// --- Siemens Structured Format ---
DATA_BLOCK "model__HS32_IW10_"
{ S7_Optimized_Access := 'TRUE' }
VERSION :
NON_RETAIN
   VAR
      W_i : ARRAY[0..31, 0..39] OF REAL;
      W_f : ARRAY[0..31, 0..39] OF REAL;
      W_g : ARRAY[0..31, 0..39] OF REAL;
      W_o : ARRAY[0..31, 0..39] OF REAL;
      R_i : ARRAY[0..31, 0..31] OF REAL;
      R_f : ARRAY[0..31, 0..31] OF REAL;
      R_g : ARRAY[0..31, 0..31] OF REAL;
      R_o : ARRAY[0..31, 0..31] OF REAL;
      B_i : ARRAY[0..31] OF REAL;
      B_f : ARRAY[0..31] OF REAL;
      B_g : ARRAY[0..31] OF REAL;
      B_o : ARRAY[0..31] OF REAL;
      FC_W : ARRAY[0..39, 0..31] OF REAL;
      FC_B : ARRAY[0..39] OF REAL;
   END_VAR
BEGIN

      W_i[0,0] := -0.10414906;
      W_i[0,1] := 0.05087908;
      W_i[0,2] := 0.03123917;
      W_i[0,3] := 0.07883381;
      W_i[0,4] := -0.04182333;
      W_i[0,5] := -0.00272775;
      W_i[0,6] := -0.10306227;
      W_i[0,7] := 0.27651954;
      W_i[0,8] := 0.07111089;
      W_i[0,9] := -0.17811616;
      W_i[0,10] := 0.00811404;
      W_i[0,11] := 0.09247471;
      W_i[0,12] := -0.06765226;
      W_i[0,13] := 0.00099094;
      W_i[0,14] := -0.00565724;
      W_i[0,15] := 0.07034151;
      W_i[0,16] := -0.03319963;
      W_i[0,17] := -0.01640407;
      W_i[0,18] := 0.00714720;
      W_i[0,19] := 0.05200255;
      W_i[0,20] := -0.10294636;
      W_i[0,21] := 0.13340643;
      W_i[0,22] := -0.48219806;
      W_i[0,23] := -0.10634176;
      W_i[0,24] := -0.78127921;
      W_i[0,25] := -0.72295207;
      W_i[0,26] := -0.21058698;
      W_i[0,27] := -0.23595250;
      W_i[0,28] := -0.07997044;
      W_i[0,29] := -0.01075801;
      W_i[0,30] := -0.32065672;
      W_i[0,31] := -0.08546381;
      W_i[0,32] := -0.13408948;
      W_i[0,33] := 0.01877546;
      W_i[0,34] := -0.84940672;
      W_i[0,35] := -0.07448237;
      W_i[0,36] := -0.02454676;
      W_i[0,37] := -0.26921397;
      W_i[0,38] := -0.07333633;
      W_i[0,39] := -0.01266416;
      W_i[1,0] := 0.29037470;
      W_i[1,1] := 0.04892659;
      W_i[1,2] := 0.02171497;
      W_i[1,3] := 0.02552549;
      W_i[1,4] := 0.01215333;
      W_i[1,5] := 0.03346634;
      W_i[1,6] := -0.03770757;
      W_i[1,7] := 0.26558429;
      W_i[1,8] := -0.11029382;
      W_i[1,9] := -0.20845115;
      W_i[1,10] := -0.01400178;
      W_i[1,11] := 0.15223934;
      W_i[1,12] := -0.13050519;
      W_i[1,13] := -0.04419332;
      W_i[1,14] := 0.00628915;
      W_i[1,15] := 0.04288426;
      W_i[1,16] := -0.00701924;
      W_i[1,17] := 0.02646778;
      W_i[1,18] := -0.00136598;
      W_i[1,19] := 0.07391773;
      W_i[1,20] := 0.03997133;
      W_i[1,21] := 0.11501998;
      W_i[1,22] := -0.30713096;
      W_i[1,23] := -0.01738190;
      W_i[1,24] := -0.39384720;
      W_i[1,25] := -0.48897827;
      W_i[1,26] := -0.01727662;
      W_i[1,27] := -0.21526198;
      W_i[1,28] := -0.00675165;
      W_i[1,29] := 0.18086264;
      W_i[1,30] := -0.21994361;
      W_i[1,31] := -0.03053124;
      W_i[1,32] := -0.17159809;
      W_i[1,33] := -0.00609811;
      W_i[1,34] := -0.71118248;
      W_i[1,35] := -0.12901427;
      W_i[1,36] := -0.05088318;
      W_i[1,37] := -0.12064310;
      W_i[1,38] := -0.03252085;
      W_i[1,39] := -0.03171032;
      W_i[2,0] := -0.00230766;
      W_i[2,1] := -0.01114088;
      W_i[2,2] := 0.00278754;
      W_i[2,3] := -0.04560725;
      W_i[2,4] := -0.00076747;
      W_i[2,5] := -0.02340589;
      W_i[2,6] := -0.09104784;
      W_i[2,7] := -0.03890763;
      W_i[2,8] := 0.02353094;
      W_i[2,9] := 0.00039863;
      W_i[2,10] := 0.01153927;
      W_i[2,11] := 0.04803184;
      W_i[2,12] := 0.08744484;
      W_i[2,13] := 0.04118077;
      W_i[2,14] := 0.02094036;
      W_i[2,15] := 0.12591685;
      W_i[2,16] := 0.01395341;
      W_i[2,17] := 0.02091648;
      W_i[2,18] := -0.04870405;
      W_i[2,19] := -0.04149374;
      W_i[2,20] := 0.10584776;
      W_i[2,21] := 0.06836145;
      W_i[2,22] := 0.01589410;
      W_i[2,23] := -0.06229543;
      W_i[2,24] := -0.27194241;
      W_i[2,25] := -0.39684960;
      W_i[2,26] := 0.03680405;
      W_i[2,27] := 0.08170957;
      W_i[2,28] := 0.08198555;
      W_i[2,29] := 0.08877461;
      W_i[2,30] := 0.25039282;
      W_i[2,31] := 0.00393842;
      W_i[2,32] := 0.15045230;
      W_i[2,33] := -0.04096574;
      W_i[2,34] := 0.44737267;
      W_i[2,35] := -0.14432395;
      W_i[2,36] := -0.04863369;
      W_i[2,37] := -0.42030501;
      W_i[2,38] := -0.05893779;
      W_i[2,39] := -0.01147668;
      W_i[3,0] := -0.11661218;
      W_i[3,1] := -0.11039881;
      W_i[3,2] := -0.09505490;
      W_i[3,3] := -0.05274161;
      W_i[3,4] := 0.13631159;
      W_i[3,5] := -0.41682443;
      W_i[3,6] := 0.34413198;
      W_i[3,7] := 0.19693865;
      W_i[3,8] := -0.37381542;
      W_i[3,9] := 0.03602328;
      W_i[3,10] := 0.32276613;
      W_i[3,11] := -0.61351973;
      W_i[3,12] := -0.15591657;
      W_i[3,13] := -0.22586936;
      W_i[3,14] := -0.00271499;
      W_i[3,15] := 0.03598518;
      W_i[3,16] := -0.04658272;
      W_i[3,17] := 0.12849101;
      W_i[3,18] := 0.14830461;
      W_i[3,19] := 0.61608970;
      W_i[3,20] := -0.01793281;
      W_i[3,21] := 0.22755618;
      W_i[3,22] := 0.04441701;
      W_i[3,23] := 0.06841668;
      W_i[3,24] := -0.42572534;
      W_i[3,25] := -0.38698140;
      W_i[3,26] := 0.11054352;
      W_i[3,27] := -0.20471475;
      W_i[3,28] := -0.03201612;
      W_i[3,29] := -0.26479176;
      W_i[3,30] := 0.02552174;
      W_i[3,31] := -0.13836773;
      W_i[3,32] := -0.11162268;
      W_i[3,33] := -0.09296755;
      W_i[3,34] := -0.26265231;
      W_i[3,35] := -0.16597824;
      W_i[3,36] := 0.03927263;
      W_i[3,37] := -0.06124702;
      W_i[3,38] := 0.16334522;
      W_i[3,39] := 0.95440286;
      W_i[4,0] := -0.09592919;
      W_i[4,1] := 0.07784065;
      W_i[4,2] := 0.01346385;
      W_i[4,3] := 0.08287931;
      W_i[4,4] := -0.42782676;
      W_i[4,5] := 0.03361791;
      W_i[4,6] := -0.15880656;
      W_i[4,7] := -0.05813188;
      W_i[4,8] := -0.01824343;
      W_i[4,9] := -0.11751872;
      W_i[4,10] := 0.14676669;
      W_i[4,11] := 0.02209505;
      W_i[4,12] := -0.00572815;
      W_i[4,13] := 0.05958780;
      W_i[4,14] := -0.02038914;
      W_i[4,15] := -0.01525941;
      W_i[4,16] := -0.03268129;
      W_i[4,17] := 0.01159987;
      W_i[4,18] := -0.02004867;
      W_i[4,19] := -0.07593681;
      W_i[4,20] := 0.05724435;
      W_i[4,21] := -0.28372633;
      W_i[4,22] := -0.11699247;
      W_i[4,23] := -0.35998097;
      W_i[4,24] := 0.26990792;
      W_i[4,25] := 0.15219623;
      W_i[4,26] := -0.08656731;
      W_i[4,27] := 0.16333446;
      W_i[4,28] := 0.13229539;
      W_i[4,29] := 0.18428297;
      W_i[4,30] := -0.18249886;
      W_i[4,31] := 0.24244712;
      W_i[4,32] := -0.00069160;
      W_i[4,33] := 0.29610279;
      W_i[4,34] := 0.03106182;
      W_i[4,35] := -0.07256878;
      W_i[4,36] := 0.03714421;
      W_i[4,37] := -0.08504521;
      W_i[4,38] := -0.01051908;
      W_i[4,39] := 0.00350483;
      W_i[5,0] := -0.05495714;
      W_i[5,1] := 0.17977138;
      W_i[5,2] := 0.04651625;
      W_i[5,3] := 0.08715992;
      W_i[5,4] := 0.10765444;
      W_i[5,5] := -0.10662776;
      W_i[5,6] := -0.04317707;
      W_i[5,7] := 0.04963618;
      W_i[5,8] := 0.00394473;
      W_i[5,9] := 0.02992170;
      W_i[5,10] := -0.02726821;
      W_i[5,11] := 0.21677773;
      W_i[5,12] := -0.15348147;
      W_i[5,13] := -0.01556183;
      W_i[5,14] := 0.01471778;
      W_i[5,15] := -0.00319904;
      W_i[5,16] := 0.06557427;
      W_i[5,17] := -0.00420085;
      W_i[5,18] := 0.00420561;
      W_i[5,19] := 0.07868493;
      W_i[5,20] := -0.17903206;
      W_i[5,21] := -0.01610633;
      W_i[5,22] := -0.42383689;
      W_i[5,23] := -0.00551023;
      W_i[5,24] := -0.38271463;
      W_i[5,25] := -0.08532900;
      W_i[5,26] := 0.03424337;
      W_i[5,27] := 0.00513940;
      W_i[5,28] := -0.12665990;
      W_i[5,29] := 0.72981369;
      W_i[5,30] := -0.61144358;
      W_i[5,31] := -0.02451378;
      W_i[5,32] := -0.15765238;
      W_i[5,33] := -0.08363440;
      W_i[5,34] := -0.17316997;
      W_i[5,35] := 0.04921770;
      W_i[5,36] := 0.03656118;
      W_i[5,37] := -0.23534429;
      W_i[5,38] := -0.03259736;
      W_i[5,39] := -0.02564295;
      W_i[6,0] := -0.07149911;
      W_i[6,1] := 0.05910936;
      W_i[6,2] := 0.02579894;
      W_i[6,3] := 0.07767012;
      W_i[6,4] := -0.02382352;
      W_i[6,5] := 0.03319338;
      W_i[6,6] := -0.03900349;
      W_i[6,7] := -0.11483924;
      W_i[6,8] := -0.07984669;
      W_i[6,9] := -0.03000957;
      W_i[6,10] := 0.04087067;
      W_i[6,11] := 0.05389729;
      W_i[6,12] := -0.15653324;
      W_i[6,13] := -0.03200754;
      W_i[6,14] := -0.00524681;
      W_i[6,15] := -0.00143958;
      W_i[6,16] := -0.01686914;
      W_i[6,17] := -0.00267206;
      W_i[6,18] := 0.03467545;
      W_i[6,19] := 0.11881366;
      W_i[6,20] := 0.15485220;
      W_i[6,21] := -0.25145912;
      W_i[6,22] := 0.02979270;
      W_i[6,23] := 0.04974350;
      W_i[6,24] := -0.06280798;
      W_i[6,25] := 0.04208164;
      W_i[6,26] := 0.06788322;
      W_i[6,27] := 0.22705127;
      W_i[6,28] := 0.07820445;
      W_i[6,29] := -0.25283822;
      W_i[6,30] := 0.02389662;
      W_i[6,31] := -0.03982587;
      W_i[6,32] := 0.08894450;
      W_i[6,33] := 0.11913013;
      W_i[6,34] := 0.21554954;
      W_i[6,35] := -0.32464555;
      W_i[6,36] := 0.02452838;
      W_i[6,37] := -0.31377190;
      W_i[6,38] := 0.00847345;
      W_i[6,39] := 0.09918413;
      W_i[7,0] := 0.02757634;
      W_i[7,1] := -0.02689262;
      W_i[7,2] := -0.02939863;
      W_i[7,3] := -0.04568179;
      W_i[7,4] := -0.09635723;
      W_i[7,5] := -0.03179899;
      W_i[7,6] := -0.12191572;
      W_i[7,7] := 0.30427256;
      W_i[7,8] := 0.21273117;
      W_i[7,9] := -0.31949016;
      W_i[7,10] := 0.01761072;
      W_i[7,11] := -0.09866854;
      W_i[7,12] := 0.10523087;
      W_i[7,13] := 0.07799035;
      W_i[7,14] := 0.07163531;
      W_i[7,15] := 0.04057769;
      W_i[7,16] := -0.03791607;
      W_i[7,17] := 0.04264954;
      W_i[7,18] := -0.09266370;
      W_i[7,19] := -0.00260587;
      W_i[7,20] := -0.03977212;
      W_i[7,21] := -0.20910311;
      W_i[7,22] := -0.00171320;
      W_i[7,23] := -0.04438376;
      W_i[7,24] := -1.20630348;
      W_i[7,25] := -0.21321478;
      W_i[7,26] := -0.06407063;
      W_i[7,27] := 0.11449858;
      W_i[7,28] := 0.03520356;
      W_i[7,29] := 0.21331252;
      W_i[7,30] := 0.21956272;
      W_i[7,31] := -0.00092769;
      W_i[7,32] := -0.11663342;
      W_i[7,33] := 0.14221379;
      W_i[7,34] := -0.10930648;
      W_i[7,35] := 0.04132334;
      W_i[7,36] := 0.05281549;
      W_i[7,37] := 0.15278573;
      W_i[7,38] := 0.15391673;
      W_i[7,39] := -0.02757900;
      W_i[8,0] := 0.05724476;
      W_i[8,1] := -0.03158160;
      W_i[8,2] := -0.11627535;
      W_i[8,3] := -0.05773278;
      W_i[8,4] := 0.07278191;
      W_i[8,5] := -0.08000189;
      W_i[8,6] := 0.02300551;
      W_i[8,7] := -0.08800174;
      W_i[8,8] := 0.20740731;
      W_i[8,9] := 0.06626759;
      W_i[8,10] := 0.04762848;
      W_i[8,11] := -0.10821844;
      W_i[8,12] := -0.12422320;
      W_i[8,13] := 0.02703045;
      W_i[8,14] := 0.00398667;
      W_i[8,15] := 0.00804039;
      W_i[8,16] := -0.14637028;
      W_i[8,17] := -0.07778820;
      W_i[8,18] := -0.09220842;
      W_i[8,19] := 0.47469196;
      W_i[8,20] := 0.02264124;
      W_i[8,21] := 0.04296339;
      W_i[8,22] := 0.04171297;
      W_i[8,23] := -0.06263759;
      W_i[8,24] := 0.27121377;
      W_i[8,25] := 0.31945908;
      W_i[8,26] := 0.14077963;
      W_i[8,27] := 0.10558233;
      W_i[8,28] := -0.00015772;
      W_i[8,29] := 0.18647811;
      W_i[8,30] := 0.11800971;
      W_i[8,31] := 0.10110309;
      W_i[8,32] := 0.01555773;
      W_i[8,33] := 0.06486533;
      W_i[8,34] := 0.31461737;
      W_i[8,35] := 0.15680584;
      W_i[8,36] := -0.01419803;
      W_i[8,37] := 0.05979521;
      W_i[8,38] := 0.22562319;
      W_i[8,39] := 0.54453236;
      W_i[9,0] := -0.45409659;
      W_i[9,1] := -0.06150096;
      W_i[9,2] := 0.49318254;
      W_i[9,3] := -0.51527238;
      W_i[9,4] := 0.12728609;
      W_i[9,5] := -0.10118011;
      W_i[9,6] := 0.29715037;
      W_i[9,7] := -0.05259424;
      W_i[9,8] := 0.01368861;
      W_i[9,9] := 0.17207454;
      W_i[9,10] := 0.11617907;
      W_i[9,11] := 0.01172454;
      W_i[9,12] := -0.30126482;
      W_i[9,13] := 0.17993747;
      W_i[9,14] := 0.08894411;
      W_i[9,15] := -0.23540320;
      W_i[9,16] := -0.15334457;
      W_i[9,17] := -0.18120950;
      W_i[9,18] := 0.09745281;
      W_i[9,19] := 0.18141954;
      W_i[9,20] := 0.10671264;
      W_i[9,21] := 0.24788895;
      W_i[9,22] := 0.13593909;
      W_i[9,23] := -0.13985786;
      W_i[9,24] := -0.24154125;
      W_i[9,25] := -0.12681547;
      W_i[9,26] := 0.20098042;
      W_i[9,27] := -0.32428232;
      W_i[9,28] := -0.32814661;
      W_i[9,29] := -0.23453857;
      W_i[9,30] := 0.12634908;
      W_i[9,31] := 0.14591648;
      W_i[9,32] := -0.03520398;
      W_i[9,33] := 0.11785780;
      W_i[9,34] := -1.13588667;
      W_i[9,35] := -0.19602355;
      W_i[9,36] := 0.09494327;
      W_i[9,37] := 0.00611658;
      W_i[9,38] := 0.19538435;
      W_i[9,39] := 0.03790567;
      W_i[10,0] := 0.08093075;
      W_i[10,1] := -0.03189079;
      W_i[10,2] := 0.00460666;
      W_i[10,3] := -0.25079808;
      W_i[10,4] := 0.12079003;
      W_i[10,5] := 0.06994910;
      W_i[10,6] := 0.01222384;
      W_i[10,7] := 0.07541763;
      W_i[10,8] := 0.05855694;
      W_i[10,9] := -0.01396475;
      W_i[10,10] := 0.02662643;
      W_i[10,11] := -0.66687572;
      W_i[10,12] := 0.49504700;
      W_i[10,13] := -0.05885675;
      W_i[10,14] := -0.11757897;
      W_i[10,15] := 0.06344132;
      W_i[10,16] := -0.02143165;
      W_i[10,17] := 0.02022251;
      W_i[10,18] := -0.03556326;
      W_i[10,19] := 0.04088999;
      W_i[10,20] := -0.08695306;
      W_i[10,21] := 0.13901219;
      W_i[10,22] := -0.04673401;
      W_i[10,23] := -0.13039219;
      W_i[10,24] := -0.02369194;
      W_i[10,25] := -0.13022855;
      W_i[10,26] := 0.15325138;
      W_i[10,27] := -0.14148274;
      W_i[10,28] := -0.10921547;
      W_i[10,29] := 0.50673056;
      W_i[10,30] := 0.16923237;
      W_i[10,31] := -0.06320494;
      W_i[10,32] := -0.08798328;
      W_i[10,33] := 0.01157838;
      W_i[10,34] := -0.41323879;
      W_i[10,35] := 0.09598303;
      W_i[10,36] := 0.02359625;
      W_i[10,37] := -0.05013705;
      W_i[10,38] := -0.02053811;
      W_i[10,39] := 1.16537046;
      W_i[11,0] := -0.13920400;
      W_i[11,1] := 0.10422801;
      W_i[11,2] := 0.05192634;
      W_i[11,3] := 0.02474182;
      W_i[11,4] := -0.11992953;
      W_i[11,5] := -0.11497844;
      W_i[11,6] := -0.06959671;
      W_i[11,7] := 0.08906282;
      W_i[11,8] := 0.00035152;
      W_i[11,9] := -0.10795452;
      W_i[11,10] := 0.02394083;
      W_i[11,11] := -0.07669503;
      W_i[11,12] := 0.15492713;
      W_i[11,13] := 0.02082890;
      W_i[11,14] := 0.01739825;
      W_i[11,15] := 0.28620026;
      W_i[11,16] := -0.05672961;
      W_i[11,17] := 0.07933230;
      W_i[11,18] := -0.19136667;
      W_i[11,19] := -0.39791319;
      W_i[11,20] := -0.13187614;
      W_i[11,21] := -0.04277104;
      W_i[11,22] := -0.11175538;
      W_i[11,23] := -0.10681376;
      W_i[11,24] := -0.71706533;
      W_i[11,25] := -0.89369446;
      W_i[11,26] := -0.04355099;
      W_i[11,27] := -0.11690557;
      W_i[11,28] := 0.17073342;
      W_i[11,29] := 0.26696113;
      W_i[11,30] := -0.03069729;
      W_i[11,31] := -0.11184800;
      W_i[11,32] := 0.15421732;
      W_i[11,33] := 0.14543033;
      W_i[11,34] := -0.00053378;
      W_i[11,35] := 0.08841224;
      W_i[11,36] := 0.00902623;
      W_i[11,37] := -0.14363292;
      W_i[11,38] := -0.02996587;
      W_i[11,39] := 0.03438438;
      W_i[12,0] := 0.02294069;
      W_i[12,1] := -0.00171102;
      W_i[12,2] := -0.00742173;
      W_i[12,3] := -0.06263760;
      W_i[12,4] := 0.01279054;
      W_i[12,5] := -0.07051820;
      W_i[12,6] := 0.03081366;
      W_i[12,7] := 0.01733820;
      W_i[12,8] := -0.01632435;
      W_i[12,9] := -0.03842505;
      W_i[12,10] := 0.11362740;
      W_i[12,11] := 0.01187946;
      W_i[12,12] := -0.19036539;
      W_i[12,13] := 0.00812287;
      W_i[12,14] := 0.00857556;
      W_i[12,15] := 0.06468427;
      W_i[12,16] := 0.01327470;
      W_i[12,17] := 0.05196055;
      W_i[12,18] := 0.00679103;
      W_i[12,19] := 0.10192532;
      W_i[12,20] := 0.01617677;
      W_i[12,21] := -0.01601717;
      W_i[12,22] := -0.22829570;
      W_i[12,23] := 0.02394662;
      W_i[12,24] := -0.15263872;
      W_i[12,25] := -0.21143152;
      W_i[12,26] := 0.02614386;
      W_i[12,27] := 0.03263390;
      W_i[12,28] := -0.02625607;
      W_i[12,29] := 0.11965574;
      W_i[12,30] := -0.15762709;
      W_i[12,31] := -0.02538990;
      W_i[12,32] := -0.08307584;
      W_i[12,33] := -0.31617489;
      W_i[12,34] := -0.47193074;
      W_i[12,35] := 0.05056112;
      W_i[12,36] := -0.02334138;
      W_i[12,37] := 0.05162949;
      W_i[12,38] := -0.00184243;
      W_i[12,39] := -0.07476960;
      W_i[13,0] := -0.05422729;
      W_i[13,1] := 0.05369066;
      W_i[13,2] := 0.19673365;
      W_i[13,3] := -0.01662629;
      W_i[13,4] := -0.25112736;
      W_i[13,5] := 0.04215603;
      W_i[13,6] := -0.01216646;
      W_i[13,7] := -0.02261561;
      W_i[13,8] := 0.06583825;
      W_i[13,9] := -0.09321744;
      W_i[13,10] := 0.09180189;
      W_i[13,11] := -0.03501062;
      W_i[13,12] := -0.05178300;
      W_i[13,13] := 0.02152647;
      W_i[13,14] := -0.00585466;
      W_i[13,15] := 0.02690242;
      W_i[13,16] := 0.05156825;
      W_i[13,17] := -0.00785884;
      W_i[13,18] := 0.03111081;
      W_i[13,19] := 0.06616246;
      W_i[13,20] := 0.37484357;
      W_i[13,21] := 0.39685732;
      W_i[13,22] := 0.24273588;
      W_i[13,23] := -0.16400047;
      W_i[13,24] := -0.48090297;
      W_i[13,25] := -0.65926820;
      W_i[13,26] := 0.00232797;
      W_i[13,27] := -0.39699012;
      W_i[13,28] := 0.19753022;
      W_i[13,29] := -0.06130902;
      W_i[13,30] := 0.28690943;
      W_i[13,31] := -0.10682096;
      W_i[13,32] := -0.20434864;
      W_i[13,33] := -0.00529929;
      W_i[13,34] := -0.08101957;
      W_i[13,35] := -0.28162447;
      W_i[13,36] := -0.00019771;
      W_i[13,37] := -0.10134698;
      W_i[13,38] := 0.08405506;
      W_i[13,39] := 0.02791081;
      W_i[14,0] := -0.00641464;
      W_i[14,1] := -0.07902622;
      W_i[14,2] := -0.00962101;
      W_i[14,3] := -0.10157780;
      W_i[14,4] := -0.20325656;
      W_i[14,5] := -0.10654134;
      W_i[14,6] := -0.17346123;
      W_i[14,7] := -0.08654054;
      W_i[14,8] := 0.04967920;
      W_i[14,9] := 0.03463001;
      W_i[14,10] := -0.01520124;
      W_i[14,11] := -0.16036510;
      W_i[14,12] := 0.11977271;
      W_i[14,13] := -0.01360948;
      W_i[14,14] := -0.02822133;
      W_i[14,15] := 0.06596331;
      W_i[14,16] := -0.03343983;
      W_i[14,17] := -0.00003674;
      W_i[14,18] := -0.01699661;
      W_i[14,19] := -0.06715041;
      W_i[14,20] := -0.00364850;
      W_i[14,21] := -0.11120961;
      W_i[14,22] := 0.13065438;
      W_i[14,23] := 0.09395862;
      W_i[14,24] := -0.16753431;
      W_i[14,25] := 0.11231579;
      W_i[14,26] := -0.08660205;
      W_i[14,27] := 0.06371113;
      W_i[14,28] := 0.22697905;
      W_i[14,29] := -0.12977916;
      W_i[14,30] := -0.05202354;
      W_i[14,31] := -0.10200743;
      W_i[14,32] := 0.23616455;
      W_i[14,33] := -0.04918646;
      W_i[14,34] := -0.09626528;
      W_i[14,35] := -0.05409024;
      W_i[14,36] := 0.06871973;
      W_i[14,37] := -0.05609881;
      W_i[14,38] := -0.02303308;
      W_i[14,39] := 0.31518012;
      W_i[15,0] := -0.09676790;
      W_i[15,1] := -0.01758914;
      W_i[15,2] := 0.04379245;
      W_i[15,3] := -0.04654387;
      W_i[15,4] := 0.01024284;
      W_i[15,5] := -0.05845871;
      W_i[15,6] := 0.00743835;
      W_i[15,7] := -0.02094029;
      W_i[15,8] := -0.09091701;
      W_i[15,9] := 0.11865507;
      W_i[15,10] := -0.01746805;
      W_i[15,11] := 0.20039460;
      W_i[15,12] := -0.12642927;
      W_i[15,13] := -0.00514105;
      W_i[15,14] := 0.03923552;
      W_i[15,15] := 0.11638938;
      W_i[15,16] := -0.07961880;
      W_i[15,17] := 0.04205161;
      W_i[15,18] := 0.25933996;
      W_i[15,19] := 0.06984173;
      W_i[15,20] := -0.05151952;
      W_i[15,21] := 0.06932238;
      W_i[15,22] := -0.07498714;
      W_i[15,23] := -0.06292155;
      W_i[15,24] := -0.49972233;
      W_i[15,25] := -0.60685724;
      W_i[15,26] := -0.05439887;
      W_i[15,27] := -0.06120267;
      W_i[15,28] := 0.00700127;
      W_i[15,29] := 0.16338313;
      W_i[15,30] := -0.16948389;
      W_i[15,31] := -0.01669374;
      W_i[15,32] := -0.25057963;
      W_i[15,33] := -0.02915098;
      W_i[15,34] := -0.68399107;
      W_i[15,35] := -0.07107162;
      W_i[15,36] := -0.05043574;
      W_i[15,37] := 0.04372098;
      W_i[15,38] := -0.25013936;
      W_i[15,39] := 0.13857038;
      W_i[16,0] := -0.02032313;
      W_i[16,1] := -0.06054825;
      W_i[16,2] := -0.05018746;
      W_i[16,3] := -0.32905868;
      W_i[16,4] := 0.03207379;
      W_i[16,5] := 0.00894374;
      W_i[16,6] := -0.07940612;
      W_i[16,7] := 0.08516731;
      W_i[16,8] := 0.17122981;
      W_i[16,9] := 0.12401859;
      W_i[16,10] := -0.00566656;
      W_i[16,11] := 0.55509824;
      W_i[16,12] := -0.12797573;
      W_i[16,13] := 0.12840185;
      W_i[16,14] := -0.00560220;
      W_i[16,15] := -0.03253403;
      W_i[16,16] := 0.09733566;
      W_i[16,17] := 0.25801903;
      W_i[16,18] := 0.11380161;
      W_i[16,19] := -0.80272037;
      W_i[16,20] := 0.04138433;
      W_i[16,21] := -0.01263740;
      W_i[16,22] := -0.04676542;
      W_i[16,23] := -0.04128587;
      W_i[16,24] := -0.09060884;
      W_i[16,25] := -0.07899155;
      W_i[16,26] := -0.06430305;
      W_i[16,27] := 0.03604764;
      W_i[16,28] := 0.00045348;
      W_i[16,29] := 0.03380001;
      W_i[16,30] := 0.00501510;
      W_i[16,31] := -0.05046950;
      W_i[16,32] := 0.04200895;
      W_i[16,33] := 0.04899995;
      W_i[16,34] := -0.29613250;
      W_i[16,35] := 0.07269148;
      W_i[16,36] := -0.01593749;
      W_i[16,37] := 0.14762485;
      W_i[16,38] := 1.97573650;
      W_i[16,39] := 0.22949235;
      W_i[17,0] := 0.08476084;
      W_i[17,1] := -0.00679670;
      W_i[17,2] := -0.22119424;
      W_i[17,3] := 0.48269364;
      W_i[17,4] := -0.11560152;
      W_i[17,5] := 0.07457293;
      W_i[17,6] := -0.09854076;
      W_i[17,7] := -0.13171072;
      W_i[17,8] := 0.10163180;
      W_i[17,9] := -0.19218649;
      W_i[17,10] := -0.30006346;
      W_i[17,11] := -0.31067795;
      W_i[17,12] := 0.37090316;
      W_i[17,13] := 0.01393779;
      W_i[17,14] := -0.04519158;
      W_i[17,15] := -0.24595827;
      W_i[17,16] := 0.13599655;
      W_i[17,17] := -0.02554221;
      W_i[17,18] := 0.07901859;
      W_i[17,19] := -0.17056887;
      W_i[17,20] := 0.17610712;
      W_i[17,21] := 0.19956675;
      W_i[17,22] := 0.26856163;
      W_i[17,23] := -0.04846491;
      W_i[17,24] := -0.35467815;
      W_i[17,25] := -0.73777598;
      W_i[17,26] := -0.00338157;
      W_i[17,27] := -0.17366287;
      W_i[17,28] := 0.04138387;
      W_i[17,29] := -0.07655122;
      W_i[17,30] := 0.23662250;
      W_i[17,31] := 0.13502227;
      W_i[17,32] := 0.06229091;
      W_i[17,33] := 0.27484414;
      W_i[17,34] := -0.36532125;
      W_i[17,35] := 0.23919977;
      W_i[17,36] := 0.03001186;
      W_i[17,37] := -0.02651701;
      W_i[17,38] := -0.10966329;
      W_i[17,39] := -0.09765702;
      W_i[18,0] := -0.01072698;
      W_i[18,1] := -0.01754156;
      W_i[18,2] := -0.06045541;
      W_i[18,3] := 0.27792412;
      W_i[18,4] := -0.10338698;
      W_i[18,5] := -0.01724318;
      W_i[18,6] := 0.05972869;
      W_i[18,7] := 0.19531298;
      W_i[18,8] := -0.04305949;
      W_i[18,9] := -0.28192112;
      W_i[18,10] := -0.01495953;
      W_i[18,11] := 0.02185066;
      W_i[18,12] := -0.03796329;
      W_i[18,13] := -0.02919699;
      W_i[18,14] := 0.01971957;
      W_i[18,15] := -0.05317892;
      W_i[18,16] := -0.01361690;
      W_i[18,17] := 0.01569653;
      W_i[18,18] := 0.04128148;
      W_i[18,19] := 0.09051883;
      W_i[18,20] := -0.08817165;
      W_i[18,21] := -0.23886830;
      W_i[18,22] := 0.05415753;
      W_i[18,23] := -0.08203930;
      W_i[18,24] := -0.56212270;
      W_i[18,25] := -0.27550292;
      W_i[18,26] := 0.14706196;
      W_i[18,27] := 0.23544437;
      W_i[18,28] := -0.12311765;
      W_i[18,29] := 0.38246083;
      W_i[18,30] := 0.04238867;
      W_i[18,31] := 0.04184147;
      W_i[18,32] := 0.02498194;
      W_i[18,33] := 0.15546310;
      W_i[18,34] := 0.17266822;
      W_i[18,35] := -0.02983394;
      W_i[18,36] := -0.04542524;
      W_i[18,37] := 0.14777139;
      W_i[18,38] := 0.05389114;
      W_i[18,39] := 0.12323732;
      W_i[19,0] := -0.04118984;
      W_i[19,1] := -0.05178985;
      W_i[19,2] := 0.01247051;
      W_i[19,3] := -0.10230274;
      W_i[19,4] := 0.06554563;
      W_i[19,5] := -0.03652082;
      W_i[19,6] := -0.01573814;
      W_i[19,7] := -0.22882380;
      W_i[19,8] := -0.01733048;
      W_i[19,9] := 0.02556017;
      W_i[19,10] := 0.12558261;
      W_i[19,11] := -0.35774660;
      W_i[19,12] := 0.35903713;
      W_i[19,13] := 0.04483967;
      W_i[19,14] := -0.07952754;
      W_i[19,15] := 0.17630176;
      W_i[19,16] := -0.09169330;
      W_i[19,17] := 0.04853094;
      W_i[19,18] := -0.29820153;
      W_i[19,19] := -0.55297935;
      W_i[19,20] := -0.11556186;
      W_i[19,21] := 0.04590010;
      W_i[19,22] := 0.06997641;
      W_i[19,23] := -0.06847610;
      W_i[19,24] := 0.93045694;
      W_i[19,25] := 0.67133164;
      W_i[19,26] := -0.02403742;
      W_i[19,27] := -0.06141511;
      W_i[19,28] := -0.09841657;
      W_i[19,29] := 0.11464830;
      W_i[19,30] := -0.05759177;
      W_i[19,31] := 0.07240915;
      W_i[19,32] := 0.02102977;
      W_i[19,33] := -0.34614226;
      W_i[19,34] := 0.13476451;
      W_i[19,35] := -0.07185577;
      W_i[19,36] := 0.01304692;
      W_i[19,37] := 0.08113710;
      W_i[19,38] := 0.08276531;
      W_i[19,39] := 0.75637919;
      W_i[20,0] := -0.04469725;
      W_i[20,1] := -0.08071249;
      W_i[20,2] := 0.08629666;
      W_i[20,3] := 0.16456899;
      W_i[20,4] := -0.14861588;
      W_i[20,5] := 0.07774629;
      W_i[20,6] := 0.01609089;
      W_i[20,7] := 0.08851504;
      W_i[20,8] := -0.01874496;
      W_i[20,9] := -0.07188217;
      W_i[20,10] := -0.08760341;
      W_i[20,11] := 0.15396829;
      W_i[20,12] := -0.03572583;
      W_i[20,13] := -0.15924498;
      W_i[20,14] := 0.01220816;
      W_i[20,15] := 0.06298544;
      W_i[20,16] := 0.03543315;
      W_i[20,17] := 0.03458498;
      W_i[20,18] := 0.00339782;
      W_i[20,19] := -0.00638131;
      W_i[20,20] := 0.00822721;
      W_i[20,21] := -0.20194745;
      W_i[20,22] := -0.05705288;
      W_i[20,23] := -0.01260474;
      W_i[20,24] := 0.03149515;
      W_i[20,25] := 0.31437719;
      W_i[20,26] := -0.05494177;
      W_i[20,27] := -0.06782775;
      W_i[20,28] := 0.00577347;
      W_i[20,29] := -0.10953689;
      W_i[20,30] := 0.15506610;
      W_i[20,31] := -0.02369651;
      W_i[20,32] := -0.15488286;
      W_i[20,33] := -0.15603501;
      W_i[20,34] := 0.06770360;
      W_i[20,35] := 0.21285588;
      W_i[20,36] := -0.13093460;
      W_i[20,37] := 0.13602462;
      W_i[20,38] := 0.03934853;
      W_i[20,39] := -0.02447999;
      W_i[21,0] := -0.27308202;
      W_i[21,1] := -0.20238131;
      W_i[21,2] := -0.01993954;
      W_i[21,3] := -0.18956275;
      W_i[21,4] := -0.74034709;
      W_i[21,5] := -0.12977587;
      W_i[21,6] := 0.02877652;
      W_i[21,7] := 0.29647660;
      W_i[21,8] := 0.30754596;
      W_i[21,9] := 0.08108461;
      W_i[21,10] := -0.09663523;
      W_i[21,11] := -0.11067218;
      W_i[21,12] := 0.18492268;
      W_i[21,13] := -0.58350122;
      W_i[21,14] := 0.00617139;
      W_i[21,15] := 0.00770027;
      W_i[21,16] := 0.02182386;
      W_i[21,17] := 0.02333870;
      W_i[21,18] := 0.82925409;
      W_i[21,19] := -0.03380872;
      W_i[21,20] := 0.35278130;
      W_i[21,21] := -0.60522830;
      W_i[21,22] := 0.05552828;
      W_i[21,23] := -0.45237646;
      W_i[21,24] := 0.01976128;
      W_i[21,25] := 0.23553391;
      W_i[21,26] := 0.32768828;
      W_i[21,27] := 0.40845692;
      W_i[21,28] := 0.41547236;
      W_i[21,29] := -0.44120485;
      W_i[21,30] := -0.12294575;
      W_i[21,31] := 0.15705259;
      W_i[21,32] := 0.01334460;
      W_i[21,33] := 0.00634381;
      W_i[21,34] := -0.05295283;
      W_i[21,35] := -0.00546547;
      W_i[21,36] := -0.01102279;
      W_i[21,37] := 0.06832597;
      W_i[21,38] := 0.33954817;
      W_i[21,39] := 0.02734024;
      W_i[22,0] := 0.05740246;
      W_i[22,1] := -0.02535794;
      W_i[22,2] := 0.03597351;
      W_i[22,3] := 0.13381189;
      W_i[22,4] := -0.02694429;
      W_i[22,5] := 0.00182078;
      W_i[22,6] := -0.06583701;
      W_i[22,7] := -0.07891550;
      W_i[22,8] := -0.16364604;
      W_i[22,9] := -0.03777923;
      W_i[22,10] := -0.10684580;
      W_i[22,11] := -0.00632763;
      W_i[22,12] := 0.17695771;
      W_i[22,13] := -0.07253629;
      W_i[22,14] := 0.08045280;
      W_i[22,15] := 0.11535356;
      W_i[22,16] := -0.09878208;
      W_i[22,17] := 0.00594875;
      W_i[22,18] := 0.02490165;
      W_i[22,19] := 0.04404743;
      W_i[22,20] := -0.02046026;
      W_i[22,21] := 0.09462272;
      W_i[22,22] := 0.05234362;
      W_i[22,23] := -0.04172071;
      W_i[22,24] := -0.16626704;
      W_i[22,25] := -0.14089724;
      W_i[22,26] := 0.12763932;
      W_i[22,27] := -0.09503621;
      W_i[22,28] := -0.01844574;
      W_i[22,29] := 0.11409646;
      W_i[22,30] := -0.15128562;
      W_i[22,31] := 0.00849273;
      W_i[22,32] := 0.04971634;
      W_i[22,33] := -0.02168483;
      W_i[22,34] := -0.15375729;
      W_i[22,35] := -0.01387732;
      W_i[22,36] := -0.02604078;
      W_i[22,37] := 0.06863436;
      W_i[22,38] := 0.19154918;
      W_i[22,39] := 0.36760291;
      W_i[23,0] := 0.34011921;
      W_i[23,1] := -0.08005925;
      W_i[23,2] := -0.62199742;
      W_i[23,3] := -0.19489965;
      W_i[23,4] := 0.03212633;
      W_i[23,5] := -0.04383887;
      W_i[23,6] := -0.19573109;
      W_i[23,7] := 0.29504162;
      W_i[23,8] := 0.19906585;
      W_i[23,9] := -0.29276019;
      W_i[23,10] := -0.14652014;
      W_i[23,11] := 0.02506773;
      W_i[23,12] := 0.28118974;
      W_i[23,13] := -0.02126036;
      W_i[23,14] := 0.03418136;
      W_i[23,15] := 0.11202367;
      W_i[23,16] := -0.05830195;
      W_i[23,17] := -0.00934210;
      W_i[23,18] := 0.14349493;
      W_i[23,19] := -0.09608027;
      W_i[23,20] := -0.07349664;
      W_i[23,21] := -0.13324311;
      W_i[23,22] := -0.01711483;
      W_i[23,23] := -0.09082118;
      W_i[23,24] := -0.53038579;
      W_i[23,25] := 0.09060598;
      W_i[23,26] := 0.10956144;
      W_i[23,27] := 0.20778604;
      W_i[23,28] := -0.07752822;
      W_i[23,29] := 0.20750724;
      W_i[23,30] := -0.04916320;
      W_i[23,31] := -0.03555354;
      W_i[23,32] := 0.22611436;
      W_i[23,33] := 0.07337805;
      W_i[23,34] := 0.06392603;
      W_i[23,35] := 0.04458339;
      W_i[23,36] := -0.01548391;
      W_i[23,37] := 0.17942379;
      W_i[23,38] := -0.05364095;
      W_i[23,39] := 0.39701992;
      W_i[24,0] := -0.11757758;
      W_i[24,1] := 0.12211614;
      W_i[24,2] := 0.01774397;
      W_i[24,3] := 0.07604476;
      W_i[24,4] := -0.13878615;
      W_i[24,5] := 0.01148156;
      W_i[24,6] := 0.02342060;
      W_i[24,7] := 0.01812497;
      W_i[24,8] := -0.07917058;
      W_i[24,9] := -0.06389529;
      W_i[24,10] := 0.09163875;
      W_i[24,11] := 0.24410519;
      W_i[24,12] := -0.11526154;
      W_i[24,13] := -0.05962858;
      W_i[24,14] := 0.00398998;
      W_i[24,15] := -0.02559417;
      W_i[24,16] := 0.00355432;
      W_i[24,17] := -0.00373959;
      W_i[24,18] := 0.03150101;
      W_i[24,19] := 0.02155573;
      W_i[24,20] := 0.03827539;
      W_i[24,21] := 0.06793781;
      W_i[24,22] := -0.10372207;
      W_i[24,23] := 0.01133421;
      W_i[24,24] := -0.62039411;
      W_i[24,25] := -0.29835266;
      W_i[24,26] := -0.03344662;
      W_i[24,27] := -0.02603021;
      W_i[24,28] := 0.15519704;
      W_i[24,29] := 0.03103866;
      W_i[24,30] := -0.18793204;
      W_i[24,31] := 0.19548637;
      W_i[24,32] := -0.05793502;
      W_i[24,33] := -0.01816287;
      W_i[24,34] := 0.27196321;
      W_i[24,35] := -0.15902427;
      W_i[24,36] := -0.09312251;
      W_i[24,37] := -0.16644843;
      W_i[24,38] := -0.06393228;
      W_i[24,39] := 0.03567641;
      W_i[25,0] := 0.06553930;
      W_i[25,1] := -0.01274281;
      W_i[25,2] := -0.05734614;
      W_i[25,3] := -0.02906677;
      W_i[25,4] := -0.02566788;
      W_i[25,5] := -0.01489288;
      W_i[25,6] := -0.02714110;
      W_i[25,7] := 0.10876387;
      W_i[25,8] := 0.13895753;
      W_i[25,9] := -0.14643434;
      W_i[25,10] := -0.02018436;
      W_i[25,11] := -0.06465659;
      W_i[25,12] := -0.00351206;
      W_i[25,13] := 0.23012245;
      W_i[25,14] := 0.00838335;
      W_i[25,15] := 0.03456668;
      W_i[25,16] := 0.00988164;
      W_i[25,17] := -0.00074405;
      W_i[25,18] := -0.01163063;
      W_i[25,19] := 0.02717012;
      W_i[25,20] := 0.08796088;
      W_i[25,21] := -0.08655845;
      W_i[25,22] := -0.11495681;
      W_i[25,23] := -0.24570324;
      W_i[25,24] := -0.12923777;
      W_i[25,25] := -0.33254570;
      W_i[25,26] := 0.06977971;
      W_i[25,27] := 0.00588068;
      W_i[25,28] := 0.11621011;
      W_i[25,29] := -0.14120518;
      W_i[25,30] := 0.09575406;
      W_i[25,31] := 0.21271861;
      W_i[25,32] := 0.02734705;
      W_i[25,33] := -0.04763836;
      W_i[25,34] := -0.12678382;
      W_i[25,35] := 0.24629676;
      W_i[25,36] := -0.03925357;
      W_i[25,37] := -0.07211839;
      W_i[25,38] := 0.05005833;
      W_i[25,39] := -0.00206914;
      W_i[26,0] := 0.14974725;
      W_i[26,1] := 0.01535374;
      W_i[26,2] := -0.00377980;
      W_i[26,3] := -0.00081873;
      W_i[26,4] := -0.02556575;
      W_i[26,5] := -0.05678970;
      W_i[26,6] := 0.01107223;
      W_i[26,7] := 0.06857505;
      W_i[26,8] := 0.01311588;
      W_i[26,9] := -0.06826829;
      W_i[26,10] := -0.01936606;
      W_i[26,11] := -0.02277778;
      W_i[26,12] := 0.06435624;
      W_i[26,13] := 0.12090050;
      W_i[26,14] := -0.03857913;
      W_i[26,15] := 0.07940848;
      W_i[26,16] := -0.02777642;
      W_i[26,17] := 0.02554570;
      W_i[26,18] := 0.96746927;
      W_i[26,19] := 0.00479337;
      W_i[26,20] := -0.16709594;
      W_i[26,21] := 0.06167128;
      W_i[26,22] := -0.01846661;
      W_i[26,23] := 0.11692691;
      W_i[26,24] := -0.67230999;
      W_i[26,25] := -0.10171942;
      W_i[26,26] := -0.19048518;
      W_i[26,27] := -0.09035464;
      W_i[26,28] := -0.27786037;
      W_i[26,29] := 0.15311232;
      W_i[26,30] := -0.02550593;
      W_i[26,31] := -0.00384994;
      W_i[26,32] := 0.00329452;
      W_i[26,33] := 0.14007947;
      W_i[26,34] := -0.00689632;
      W_i[26,35] := 0.06500275;
      W_i[26,36] := -0.02411593;
      W_i[26,37] := -0.02727453;
      W_i[26,38] := 0.02548786;
      W_i[26,39] := -0.08337803;
      W_i[27,0] := 0.03984790;
      W_i[27,1] := 0.21849002;
      W_i[27,2] := 0.05760974;
      W_i[27,3] := -0.11054909;
      W_i[27,4] := 0.33313975;
      W_i[27,5] := -0.02336766;
      W_i[27,6] := -0.02719049;
      W_i[27,7] := 0.01098777;
      W_i[27,8] := 0.08218465;
      W_i[27,9] := -0.07680017;
      W_i[27,10] := -0.02052933;
      W_i[27,11] := 0.21041244;
      W_i[27,12] := -0.08520587;
      W_i[27,13] := -0.01218674;
      W_i[27,14] := 0.00151642;
      W_i[27,15] := -0.03672955;
      W_i[27,16] := 0.00260637;
      W_i[27,17] := 0.03174125;
      W_i[27,18] := -0.00094590;
      W_i[27,19] := 0.12404852;
      W_i[27,20] := 0.15310773;
      W_i[27,21] := 0.45289695;
      W_i[27,22] := -0.13904996;
      W_i[27,23] := 0.29992726;
      W_i[27,24] := 0.20153445;
      W_i[27,25] := 0.16071327;
      W_i[27,26] := 0.00996626;
      W_i[27,27] := -0.11496834;
      W_i[27,28] := -0.09930631;
      W_i[27,29] := -0.11272246;
      W_i[27,30] := -0.07931732;
      W_i[27,31] := -0.14272773;
      W_i[27,32] := -0.12526496;
      W_i[27,33] := 0.23920020;
      W_i[27,34] := 0.08852232;
      W_i[27,35] := -0.20820323;
      W_i[27,36] := 0.14521699;
      W_i[27,37] := -0.19162981;
      W_i[27,38] := 0.06865614;
      W_i[27,39] := 0.03677582;
      W_i[28,0] := 0.04997422;
      W_i[28,1] := -0.02473807;
      W_i[28,2] := -0.07641364;
      W_i[28,3] := -0.02846665;
      W_i[28,4] := -0.02600389;
      W_i[28,5] := -0.01425854;
      W_i[28,6] := 0.02516984;
      W_i[28,7] := 0.56388134;
      W_i[28,8] := 0.07125960;
      W_i[28,9] := -0.46600685;
      W_i[28,10] := -0.06418919;
      W_i[28,11] := 0.24955207;
      W_i[28,12] := -0.09087826;
      W_i[28,13] := -0.01976197;
      W_i[28,14] := 0.05677757;
      W_i[28,15] := 0.00407595;
      W_i[28,16] := -0.04238077;
      W_i[28,17] := 0.02735240;
      W_i[28,18] := -0.01160267;
      W_i[28,19] := 0.05880483;
      W_i[28,20] := 0.03925076;
      W_i[28,21] := -0.03376312;
      W_i[28,22] := 0.34712178;
      W_i[28,23] := -0.13167503;
      W_i[28,24] := -0.31470102;
      W_i[28,25] := -0.34818864;
      W_i[28,26] := -0.01199263;
      W_i[28,27] := -0.11349533;
      W_i[28,28] := -0.07639381;
      W_i[28,29] := 0.20393789;
      W_i[28,30] := 0.16922227;
      W_i[28,31] := 0.07852437;
      W_i[28,32] := 0.09054390;
      W_i[28,33] := 0.02347955;
      W_i[28,34] := -0.12864402;
      W_i[28,35] := 0.08776911;
      W_i[28,36] := -0.04564888;
      W_i[28,37] := 0.18246073;
      W_i[28,38] := -0.06260310;
      W_i[28,39] := -0.05331490;
      W_i[29,0] := 0.08882844;
      W_i[29,1] := 0.32015932;
      W_i[29,2] := 0.04887038;
      W_i[29,3] := 0.79705662;
      W_i[29,4] := -0.43447351;
      W_i[29,5] := 1.44478238;
      W_i[29,6] := 0.07902924;
      W_i[29,7] := 0.19413471;
      W_i[29,8] := -0.36958483;
      W_i[29,9] := -0.03968559;
      W_i[29,10] := 1.24356449;
      W_i[29,11] := -0.17663658;
      W_i[29,12] := 0.07064923;
      W_i[29,13] := 0.35462961;
      W_i[29,14] := 0.29002810;
      W_i[29,15] := -0.05374714;
      W_i[29,16] := 0.07444047;
      W_i[29,17] := -0.01712505;
      W_i[29,18] := 0.05375896;
      W_i[29,19] := 0.05255156;
      W_i[29,20] := -0.26016051;
      W_i[29,21] := 0.21038072;
      W_i[29,22] := -0.13402782;
      W_i[29,23] := -0.00425044;
      W_i[29,24] := 0.23636276;
      W_i[29,25] := 0.06888721;
      W_i[29,26] := -0.33938631;
      W_i[29,27] := 0.19366139;
      W_i[29,28] := 0.20567542;
      W_i[29,29] := -0.52033865;
      W_i[29,30] := -0.03867699;
      W_i[29,31] := 0.10740498;
      W_i[29,32] := 0.20093004;
      W_i[29,33] := -0.13926220;
      W_i[29,34] := -0.20935415;
      W_i[29,35] := -0.08176949;
      W_i[29,36] := -0.02408343;
      W_i[29,37] := -0.01565829;
      W_i[29,38] := 0.12726374;
      W_i[29,39] := -0.13060087;
      W_i[30,0] := -0.02755127;
      W_i[30,1] := 0.09685323;
      W_i[30,2] := 0.03178624;
      W_i[30,3] := -0.81790167;
      W_i[30,4] := -0.09512409;
      W_i[30,5] := 0.15579517;
      W_i[30,6] := -0.35025209;
      W_i[30,7] := 0.38375428;
      W_i[30,8] := 0.26148325;
      W_i[30,9] := 0.34516314;
      W_i[30,10] := -0.01904444;
      W_i[30,11] := 0.37324813;
      W_i[30,12] := 0.40989080;
      W_i[30,13] := -0.17973639;
      W_i[30,14] := 0.08796087;
      W_i[30,15] := -0.37388811;
      W_i[30,16] := -0.33972195;
      W_i[30,17] := 0.12072887;
      W_i[30,18] := 0.34597054;
      W_i[30,19] := -0.28983161;
      W_i[30,20] := -0.23207320;
      W_i[30,21] := 0.06022831;
      W_i[30,22] := 0.05972358;
      W_i[30,23] := -0.04532034;
      W_i[30,24] := -0.14049536;
      W_i[30,25] := -0.38210469;
      W_i[30,26] := 0.08971685;
      W_i[30,27] := 0.24931312;
      W_i[30,28] := 0.19635232;
      W_i[30,29] := -0.14961366;
      W_i[30,30] := -0.05470202;
      W_i[30,31] := -0.48900372;
      W_i[30,32] := 0.09259362;
      W_i[30,33] := 0.20682643;
      W_i[30,34] := -0.04097397;
      W_i[30,35] := 0.06544437;
      W_i[30,36] := -0.04607715;
      W_i[30,37] := 0.17287830;
      W_i[30,38] := 0.03883581;
      W_i[30,39] := 0.92405421;
      W_i[31,0] := 0.06235947;
      W_i[31,1] := 0.02632081;
      W_i[31,2] := -0.07524684;
      W_i[31,3] := 0.07101320;
      W_i[31,4] := -0.04651680;
      W_i[31,5] := -0.14746962;
      W_i[31,6] := 0.02125872;
      W_i[31,7] := -0.00950570;
      W_i[31,8] := 0.03748577;
      W_i[31,9] := 0.03555158;
      W_i[31,10] := 0.06589699;
      W_i[31,11] := -0.05763013;
      W_i[31,12] := 0.07570665;
      W_i[31,13] := -0.04154845;
      W_i[31,14] := -0.02712471;
      W_i[31,15] := 0.06376572;
      W_i[31,16] := -0.00796349;
      W_i[31,17] := 0.04039724;
      W_i[31,18] := -0.11584114;
      W_i[31,19] := -0.05020886;
      W_i[31,20] := 0.03928347;
      W_i[31,21] := -0.01710388;
      W_i[31,22] := -0.28104821;
      W_i[31,23] := -0.05397440;
      W_i[31,24] := 0.48354673;
      W_i[31,25] := 0.31770724;
      W_i[31,26] := 0.06595083;
      W_i[31,27] := 0.11622475;
      W_i[31,28] := -0.07772405;
      W_i[31,29] := -0.14774537;
      W_i[31,30] := -0.29682872;
      W_i[31,31] := 0.06653072;
      W_i[31,32] := -0.34515795;
      W_i[31,33] := 0.08919729;
      W_i[31,34] := -0.64831716;
      W_i[31,35] := -0.01203564;
      W_i[31,36] := -0.03006219;
      W_i[31,37] := -0.11853622;
      W_i[31,38] := 0.16422081;
      W_i[31,39] := -0.08044879;
      W_f[0,0] := -0.31087899;
      W_f[0,1] := -0.01642113;
      W_f[0,2] := -0.05293131;
      W_f[0,3] := 0.66893762;
      W_f[0,4] := -0.03667010;
      W_f[0,5] := 0.08088744;
      W_f[0,6] := -0.00525074;
      W_f[0,7] := -0.11897004;
      W_f[0,8] := -0.30270699;
      W_f[0,9] := -0.03488322;
      W_f[0,10] := 0.12175234;
      W_f[0,11] := -0.14962083;
      W_f[0,12] := 0.08034969;
      W_f[0,13] := -0.01022713;
      W_f[0,14] := 0.07079872;
      W_f[0,15] := 0.19599691;
      W_f[0,16] := -0.06211102;
      W_f[0,17] := 0.03387687;
      W_f[0,18] := -0.14573583;
      W_f[0,19] := -0.50526828;
      W_f[0,20] := -0.15081304;
      W_f[0,21] := 0.03080749;
      W_f[0,22] := -0.18689804;
      W_f[0,23] := -0.02657967;
      W_f[0,24] := 0.06952211;
      W_f[0,25] := 0.26585165;
      W_f[0,26] := -0.17459789;
      W_f[0,27] := -0.17294747;
      W_f[0,28] := 0.08707468;
      W_f[0,29] := -0.23360135;
      W_f[0,30] := -0.14734191;
      W_f[0,31] := -0.22190665;
      W_f[0,32] := -0.09349395;
      W_f[0,33] := 0.15165256;
      W_f[0,34] := -0.04947405;
      W_f[0,35] := -0.02839872;
      W_f[0,36] := -0.05069589;
      W_f[0,37] := 0.00841171;
      W_f[0,38] := 0.16808885;
      W_f[0,39] := 0.02463646;
      W_f[1,0] := 0.10309164;
      W_f[1,1] := -0.04881949;
      W_f[1,2] := -0.10869338;
      W_f[1,3] := -0.13907683;
      W_f[1,4] := -0.00155219;
      W_f[1,5] := 0.05452135;
      W_f[1,6] := -0.14117274;
      W_f[1,7] := 0.25483197;
      W_f[1,8] := -0.79242134;
      W_f[1,9] := 0.24828286;
      W_f[1,10] := 0.05196439;
      W_f[1,11] := -0.06068465;
      W_f[1,12] := -0.11384691;
      W_f[1,13] := 0.04661793;
      W_f[1,14] := 0.01614169;
      W_f[1,15] := 0.08351095;
      W_f[1,16] := 0.00189460;
      W_f[1,17] := -0.01351131;
      W_f[1,18] := 0.03005760;
      W_f[1,19] := -0.04696568;
      W_f[1,20] := -0.13451375;
      W_f[1,21] := -0.16530699;
      W_f[1,22] := 0.09706016;
      W_f[1,23] := -0.03441914;
      W_f[1,24] := -0.11357319;
      W_f[1,25] := -0.33677301;
      W_f[1,26] := 0.01804815;
      W_f[1,27] := 0.34698701;
      W_f[1,28] := 0.14250018;
      W_f[1,29] := -0.20205298;
      W_f[1,30] := 0.02922465;
      W_f[1,31] := -0.09243742;
      W_f[1,32] := 0.10971645;
      W_f[1,33] := 0.09958702;
      W_f[1,34] := -0.26081911;
      W_f[1,35] := 0.10740673;
      W_f[1,36] := 0.00407260;
      W_f[1,37] := 0.17656624;
      W_f[1,38] := -0.03367357;
      W_f[1,39] := 0.02457568;
      W_f[2,0] := 0.04323589;
      W_f[2,1] := 0.13192843;
      W_f[2,2] := -0.21908981;
      W_f[2,3] := 0.24549797;
      W_f[2,4] := -0.00847173;
      W_f[2,5] := 0.16698520;
      W_f[2,6] := 0.01734499;
      W_f[2,7] := -0.08778935;
      W_f[2,8] := -0.00173907;
      W_f[2,9] := -0.01823302;
      W_f[2,10] := -0.08939531;
      W_f[2,11] := -0.03136157;
      W_f[2,12] := -0.03248491;
      W_f[2,13] := -0.04673289;
      W_f[2,14] := -0.13506411;
      W_f[2,15] := 0.01751995;
      W_f[2,16] := 0.01984352;
      W_f[2,17] := -0.26506427;
      W_f[2,18] := -0.11390819;
      W_f[2,19] := -0.17862549;
      W_f[2,20] := -0.08476356;
      W_f[2,21] := -0.18915263;
      W_f[2,22] := 0.31209731;
      W_f[2,23] := -0.10005450;
      W_f[2,24] := 1.96645951;
      W_f[2,25] := 1.80065846;
      W_f[2,26] := -0.24080534;
      W_f[2,27] := -0.01604153;
      W_f[2,28] := -0.14632852;
      W_f[2,29] := 0.14218122;
      W_f[2,30] := 0.16648325;
      W_f[2,31] := -0.06772677;
      W_f[2,32] := 0.12971835;
      W_f[2,33] := -0.14491805;
      W_f[2,34] := 1.91479826;
      W_f[2,35] := 0.17752430;
      W_f[2,36] := 0.08425347;
      W_f[2,37] := 0.19955210;
      W_f[2,38] := 0.05383398;
      W_f[2,39] := 0.08709066;
      W_f[3,0] := -0.01027072;
      W_f[3,1] := -0.13289191;
      W_f[3,2] := -0.29553708;
      W_f[3,3] := -0.22534584;
      W_f[3,4] := -0.05643518;
      W_f[3,5] := -0.30458441;
      W_f[3,6] := 0.27409679;
      W_f[3,7] := 0.36308911;
      W_f[3,8] := -0.56274730;
      W_f[3,9] := 0.26823741;
      W_f[3,10] := 0.40326482;
      W_f[3,11] := -0.26395056;
      W_f[3,12] := -0.25299162;
      W_f[3,13] := -0.24141958;
      W_f[3,14] := -0.40557349;
      W_f[3,15] := -0.02736670;
      W_f[3,16] := 0.15541768;
      W_f[3,17] := 0.56699401;
      W_f[3,18] := 0.13678457;
      W_f[3,19] := 0.94581527;
      W_f[3,20] := 0.06098880;
      W_f[3,21] := 0.29283985;
      W_f[3,22] := -0.07756051;
      W_f[3,23] := 0.24745731;
      W_f[3,24] := -0.76781762;
      W_f[3,25] := -0.96796930;
      W_f[3,26] := 0.07189273;
      W_f[3,27] := -0.23268655;
      W_f[3,28] := -0.02444601;
      W_f[3,29] := -0.22892441;
      W_f[3,30] := 0.06516360;
      W_f[3,31] := -0.07039160;
      W_f[3,32] := -0.10594028;
      W_f[3,33] := 0.07055102;
      W_f[3,34] := -0.87469828;
      W_f[3,35] := -0.25842682;
      W_f[3,36] := -0.03514070;
      W_f[3,37] := -0.21496108;
      W_f[3,38] := -0.02638236;
      W_f[3,39] := 1.49122667;
      W_f[4,0] := -0.16676553;
      W_f[4,1] := 0.01176612;
      W_f[4,2] := 0.30374086;
      W_f[4,3] := -0.16652118;
      W_f[4,4] := 0.23176482;
      W_f[4,5] := -0.01160300;
      W_f[4,6] := -0.04741637;
      W_f[4,7] := -0.23041104;
      W_f[4,8] := -0.03371903;
      W_f[4,9] := -0.20603402;
      W_f[4,10] := 0.41277230;
      W_f[4,11] := -0.09772890;
      W_f[4,12] := -0.09781816;
      W_f[4,13] := -0.48620504;
      W_f[4,14] := 0.03265836;
      W_f[4,15] := 0.09504089;
      W_f[4,16] := 0.02240698;
      W_f[4,17] := -0.02351275;
      W_f[4,18] := -0.04697651;
      W_f[4,19] := -0.02782584;
      W_f[4,20] := 0.15254140;
      W_f[4,21] := 0.27034724;
      W_f[4,22] := 0.18237519;
      W_f[4,23] := 0.88770163;
      W_f[4,24] := -1.48963082;
      W_f[4,25] := -0.61802244;
      W_f[4,26] := -0.16299020;
      W_f[4,27] := 0.00145082;
      W_f[4,28] := 0.02346218;
      W_f[4,29] := 0.41588426;
      W_f[4,30] := 0.14504674;
      W_f[4,31] := -0.02832477;
      W_f[4,32] := 0.09136293;
      W_f[4,33] := 0.18777427;
      W_f[4,34] := -0.02872102;
      W_f[4,35] := 0.28219485;
      W_f[4,36] := -0.09533136;
      W_f[4,37] := 0.28597316;
      W_f[4,38] := 0.05682571;
      W_f[4,39] := -0.04898876;
      W_f[5,0] := 0.10161789;
      W_f[5,1] := 0.33646879;
      W_f[5,2] := -0.25958875;
      W_f[5,3] := 0.00375745;
      W_f[5,4] := -0.07752838;
      W_f[5,5] := 0.06933056;
      W_f[5,6] := -0.05768353;
      W_f[5,7] := 0.12656887;
      W_f[5,8] := 0.03442563;
      W_f[5,9] := 0.06407838;
      W_f[5,10] := -0.22720173;
      W_f[5,11] := -0.34898725;
      W_f[5,12] := -0.31888863;
      W_f[5,13] := 0.19793886;
      W_f[5,14] := -0.16154088;
      W_f[5,15] := -0.13792320;
      W_f[5,16] := -0.01594777;
      W_f[5,17] := -0.23877142;
      W_f[5,18] := -0.14457780;
      W_f[5,19] := -0.09563981;
      W_f[5,20] := -0.08250628;
      W_f[5,21] := -0.13814838;
      W_f[5,22] := 0.28552571;
      W_f[5,23] := -0.13627250;
      W_f[5,24] := 1.85639691;
      W_f[5,25] := 1.62530053;
      W_f[5,26] := -0.26891711;
      W_f[5,27] := 0.25958720;
      W_f[5,28] := 0.07219080;
      W_f[5,29] := 0.04693827;
      W_f[5,30] := 0.15581432;
      W_f[5,31] := -0.08130801;
      W_f[5,32] := 0.16866112;
      W_f[5,33] := 0.15934782;
      W_f[5,34] := 0.33171639;
      W_f[5,35] := 0.26894227;
      W_f[5,36] := 0.08339840;
      W_f[5,37] := 0.25810409;
      W_f[5,38] := -0.11701190;
      W_f[5,39] := 0.35744828;
      W_f[6,0] := -0.08564612;
      W_f[6,1] := -0.01010586;
      W_f[6,2] := 0.00021706;
      W_f[6,3] := 0.29889423;
      W_f[6,4] := 0.06283986;
      W_f[6,5] := 0.02952686;
      W_f[6,6] := 0.07751884;
      W_f[6,7] := 0.10801284;
      W_f[6,8] := -0.09512047;
      W_f[6,9] := -0.26914835;
      W_f[6,10] := -0.09744307;
      W_f[6,11] := 0.09159194;
      W_f[6,12] := 0.09488866;
      W_f[6,13] := 0.21247515;
      W_f[6,14] := -0.06295278;
      W_f[6,15] := -0.17113642;
      W_f[6,16] := -0.16463363;
      W_f[6,17] := -0.01280473;
      W_f[6,18] := -0.06927878;
      W_f[6,19] := -0.16039206;
      W_f[6,20] := -0.12198957;
      W_f[6,21] := -0.19269027;
      W_f[6,22] := 0.16312140;
      W_f[6,23] := -0.12505320;
      W_f[6,24] := 1.21596706;
      W_f[6,25] := 1.20752811;
      W_f[6,26] := -0.13087872;
      W_f[6,27] := 0.23864806;
      W_f[6,28] := -0.01269126;
      W_f[6,29] := -0.14394394;
      W_f[6,30] := 0.04508471;
      W_f[6,31] := -0.16830671;
      W_f[6,32] := 0.03094850;
      W_f[6,33] := -0.05589656;
      W_f[6,34] := 1.26290429;
      W_f[6,35] := 0.08352999;
      W_f[6,36] := 0.09383605;
      W_f[6,37] := -0.05050451;
      W_f[6,38] := 0.00890886;
      W_f[6,39] := 0.26133564;
      W_f[7,0] := -0.00092446;
      W_f[7,1] := 0.01561106;
      W_f[7,2] := -0.02553785;
      W_f[7,3] := -0.14090878;
      W_f[7,4] := 0.08901426;
      W_f[7,5] := 0.03557171;
      W_f[7,6] := 0.06185073;
      W_f[7,7] := -0.28613383;
      W_f[7,8] := 0.15983410;
      W_f[7,9] := -0.01696404;
      W_f[7,10] := -0.05231231;
      W_f[7,11] := -0.02403463;
      W_f[7,12] := 0.05044018;
      W_f[7,13] := 0.08024644;
      W_f[7,14] := -0.12023684;
      W_f[7,15] := -0.20359105;
      W_f[7,16] := 0.06390475;
      W_f[7,17] := 0.06704516;
      W_f[7,18] := 0.05190700;
      W_f[7,19] := -0.05760851;
      W_f[7,20] := 0.14534676;
      W_f[7,21] := 0.07754763;
      W_f[7,22] := -0.05249873;
      W_f[7,23] := -0.08908582;
      W_f[7,24] := -1.17519712;
      W_f[7,25] := -0.01054784;
      W_f[7,26] := 0.08837862;
      W_f[7,27] := 0.09662017;
      W_f[7,28] := -0.01325287;
      W_f[7,29] := 0.36907411;
      W_f[7,30] := 0.00725335;
      W_f[7,31] := 0.00701370;
      W_f[7,32] := 0.22163008;
      W_f[7,33] := 0.01882857;
      W_f[7,34] := 0.01451610;
      W_f[7,35] := 0.01938067;
      W_f[7,36] := 0.30278206;
      W_f[7,37] := -0.00846053;
      W_f[7,38] := -0.07525756;
      W_f[7,39] := 0.17255557;
      W_f[8,0] := 0.13039361;
      W_f[8,1] := 0.03875940;
      W_f[8,2] := -0.14218862;
      W_f[8,3] := -0.12328728;
      W_f[8,4] := -0.13652091;
      W_f[8,5] := -0.06255179;
      W_f[8,6] := -0.02927461;
      W_f[8,7] := 0.19883646;
      W_f[8,8] := -0.06549737;
      W_f[8,9] := -0.07066058;
      W_f[8,10] := 0.09409045;
      W_f[8,11] := -0.09675022;
      W_f[8,12] := 0.08247706;
      W_f[8,13] := -0.00751409;
      W_f[8,14] := 0.14233628;
      W_f[8,15] := -0.13774353;
      W_f[8,16] := 0.45766559;
      W_f[8,17] := -0.22157320;
      W_f[8,18] := 0.12065386;
      W_f[8,19] := 0.40282315;
      W_f[8,20] := 0.00461689;
      W_f[8,21] := -0.29562521;
      W_f[8,22] := -0.25563526;
      W_f[8,23] := -0.08439282;
      W_f[8,24] := -0.29703891;
      W_f[8,25] := -0.47947335;
      W_f[8,26] := -0.10692279;
      W_f[8,27] := 0.13302235;
      W_f[8,28] := 0.05997621;
      W_f[8,29] := -0.14819831;
      W_f[8,30] := -0.29963812;
      W_f[8,31] := 0.19096144;
      W_f[8,32] := -0.00359912;
      W_f[8,33] := -0.02025813;
      W_f[8,34] := -0.42184028;
      W_f[8,35] := -0.05010535;
      W_f[8,36] := -0.06069054;
      W_f[8,37] := 0.08100205;
      W_f[8,38] := -0.11007889;
      W_f[8,39] := -0.07116549;
      W_f[9,0] := -0.60376549;
      W_f[9,1] := -0.07527776;
      W_f[9,2] := 0.65037543;
      W_f[9,3] := -0.79024035;
      W_f[9,4] := -0.00867934;
      W_f[9,5] := -0.17809720;
      W_f[9,6] := 0.45782736;
      W_f[9,7] := -0.10163368;
      W_f[9,8] := -0.02632706;
      W_f[9,9] := 0.34545535;
      W_f[9,10] := 0.15282393;
      W_f[9,11] := -0.18461947;
      W_f[9,12] := -0.07619403;
      W_f[9,13] := -0.03189026;
      W_f[9,14] := 0.23177136;
      W_f[9,15] := -0.31177118;
      W_f[9,16] := -0.32775646;
      W_f[9,17] := -0.40041563;
      W_f[9,18] := 0.01072187;
      W_f[9,19] := 0.22459725;
      W_f[9,20] := 0.25021112;
      W_f[9,21] := 0.33965012;
      W_f[9,22] := -0.08007015;
      W_f[9,23] := 0.13231230;
      W_f[9,24] := -1.19737792;
      W_f[9,25] := -1.32460630;
      W_f[9,26] := 0.28357303;
      W_f[9,27] := -0.46705270;
      W_f[9,28] := -0.18736649;
      W_f[9,29] := 0.40982211;
      W_f[9,30] := -0.22468941;
      W_f[9,31] := 0.28924128;
      W_f[9,32] := -0.00599906;
      W_f[9,33] := 0.41959521;
      W_f[9,34] := 0.24919745;
      W_f[9,35] := -0.06532279;
      W_f[9,36] := 0.14215249;
      W_f[9,37] := -0.41311255;
      W_f[9,38] := 0.26410219;
      W_f[9,39] := 0.02192991;
      W_f[10,0] := 0.03587366;
      W_f[10,1] := -0.24204130;
      W_f[10,2] := 0.52407765;
      W_f[10,3] := -0.22102664;
      W_f[10,4] := -0.46720135;
      W_f[10,5] := 0.20158556;
      W_f[10,6] := 0.00767251;
      W_f[10,7] := -0.12470087;
      W_f[10,8] := 0.24142028;
      W_f[10,9] := -0.02993156;
      W_f[10,10] := -0.04576334;
      W_f[10,11] := -0.38690701;
      W_f[10,12] := 0.04477939;
      W_f[10,13] := -0.77852243;
      W_f[10,14] := -0.26673898;
      W_f[10,15] := 0.07689933;
      W_f[10,16] := -0.01653192;
      W_f[10,17] := 0.68285608;
      W_f[10,18] := -0.24064317;
      W_f[10,19] := 0.33158067;
      W_f[10,20] := -0.13776232;
      W_f[10,21] := -0.29165766;
      W_f[10,22] := 0.01264445;
      W_f[10,23] := -0.35607785;
      W_f[10,24] := 0.33992043;
      W_f[10,25] := 0.21914977;
      W_f[10,26] := 0.51194930;
      W_f[10,27] := -0.00456741;
      W_f[10,28] := 0.17721994;
      W_f[10,29] := 0.74289769;
      W_f[10,30] := -0.04158311;
      W_f[10,31] := 0.09101373;
      W_f[10,32] := -0.06729753;
      W_f[10,33] := 0.24987862;
      W_f[10,34] := 0.14726782;
      W_f[10,35] := -0.13635999;
      W_f[10,36] := -0.14212158;
      W_f[10,37] := -0.07058483;
      W_f[10,38] := 0.01411692;
      W_f[10,39] := 0.56364352;
      W_f[11,0] := -0.22232492;
      W_f[11,1] := 0.08132177;
      W_f[11,2] := -0.00592427;
      W_f[11,3] := -0.11568832;
      W_f[11,4] := -0.12797070;
      W_f[11,5] := 0.03546190;
      W_f[11,6] := 0.01878986;
      W_f[11,7] := -0.05625603;
      W_f[11,8] := 0.04217658;
      W_f[11,9] := 0.17259139;
      W_f[11,10] := -0.04498037;
      W_f[11,11] := -0.02322526;
      W_f[11,12] := 0.14480929;
      W_f[11,13] := -0.32121664;
      W_f[11,14] := -0.02877496;
      W_f[11,15] := 0.11884735;
      W_f[11,16] := -0.04417537;
      W_f[11,17] := -0.08211292;
      W_f[11,18] := -0.13818231;
      W_f[11,19] := -0.26458630;
      W_f[11,20] := -0.01089744;
      W_f[11,21] := 0.13274096;
      W_f[11,22] := -0.31027782;
      W_f[11,23] := 0.12532504;
      W_f[11,24] := -0.37777963;
      W_f[11,25] := -0.33644673;
      W_f[11,26] := -0.18400931;
      W_f[11,27] := -0.09935941;
      W_f[11,28] := 0.25673282;
      W_f[11,29] := 0.19466680;
      W_f[11,30] := -0.08646595;
      W_f[11,31] := -0.26992974;
      W_f[11,32] := -0.22119014;
      W_f[11,33] := 0.05552119;
      W_f[11,34] := 0.53751451;
      W_f[11,35] := -0.05215225;
      W_f[11,36] := 0.17789726;
      W_f[11,37] := -0.10156243;
      W_f[11,38] := -0.08626166;
      W_f[11,39] := 0.00613706;
      W_f[12,0] := 0.12016000;
      W_f[12,1] := 0.06109352;
      W_f[12,2] := -0.00014051;
      W_f[12,3] := -0.05928172;
      W_f[12,4] := -0.07623916;
      W_f[12,5] := 0.13642152;
      W_f[12,6] := -0.05664429;
      W_f[12,7] := -0.08431683;
      W_f[12,8] := -0.32728219;
      W_f[12,9] := 0.15672508;
      W_f[12,10] := -0.16274835;
      W_f[12,11] := -0.12257247;
      W_f[12,12] := -0.15561372;
      W_f[12,13] := 0.00125519;
      W_f[12,14] := 0.08071522;
      W_f[12,15] := -0.35842443;
      W_f[12,16] := -0.07716373;
      W_f[12,17] := 0.04766509;
      W_f[12,18] := 0.16450228;
      W_f[12,19] := -0.10028939;
      W_f[12,20] := -0.15282200;
      W_f[12,21] := -0.10721114;
      W_f[12,22] := -0.09602195;
      W_f[12,23] := -0.06921818;
      W_f[12,24] := 0.19129385;
      W_f[12,25] := 0.15350267;
      W_f[12,26] := -0.04103877;
      W_f[12,27] := 0.15455210;
      W_f[12,28] := -0.07642417;
      W_f[12,29] := -0.03135392;
      W_f[12,30] := 0.05042620;
      W_f[12,31] := -0.01565356;
      W_f[12,32] := -0.20334800;
      W_f[12,33] := -0.01682312;
      W_f[12,34] := -0.32919499;
      W_f[12,35] := 0.03103065;
      W_f[12,36] := -0.00876824;
      W_f[12,37] := 0.11396129;
      W_f[12,38] := 0.02205051;
      W_f[12,39] := -0.14877743;
      W_f[13,0] := -0.19990104;
      W_f[13,1] := -0.02693051;
      W_f[13,2] := -0.13122162;
      W_f[13,3] := 0.10237550;
      W_f[13,4] := 0.36373648;
      W_f[13,5] := 0.23774576;
      W_f[13,6] := 0.01520107;
      W_f[13,7] := 0.08032186;
      W_f[13,8] := 0.05583947;
      W_f[13,9] := -0.03193354;
      W_f[13,10] := -0.11794095;
      W_f[13,11] := 0.00260050;
      W_f[13,12] := -0.20683330;
      W_f[13,13] := 0.08716767;
      W_f[13,14] := -0.05809921;
      W_f[13,15] := -0.25644478;
      W_f[13,16] := -0.19208577;
      W_f[13,17] := 0.00163484;
      W_f[13,18] := -0.11728875;
      W_f[13,19] := -0.21184893;
      W_f[13,20] := -0.50744122;
      W_f[13,21] := -0.37115288;
      W_f[13,22] := 0.10131563;
      W_f[13,23] := -0.09726343;
      W_f[13,24] := 2.36166120;
      W_f[13,25] := 2.21571159;
      W_f[13,26] := -0.19924188;
      W_f[13,27] := -0.02779500;
      W_f[13,28] := 0.10948692;
      W_f[13,29] := 0.04464628;
      W_f[13,30] := 0.15166532;
      W_f[13,31] := -0.43087655;
      W_f[13,32] := 0.19548319;
      W_f[13,33] := -0.02293641;
      W_f[13,34] := 2.17658234;
      W_f[13,35] := 0.24361719;
      W_f[13,36] := -0.02843551;
      W_f[13,37] := 0.30465350;
      W_f[13,38] := 0.04337556;
      W_f[13,39] := -0.00615159;
      W_f[14,0] := -0.12647852;
      W_f[14,1] := 0.04486486;
      W_f[14,2] := 0.30913579;
      W_f[14,3] := -0.47282296;
      W_f[14,4] := -0.72544724;
      W_f[14,5] := -0.45098802;
      W_f[14,6] := -0.52586150;
      W_f[14,7] := 0.01496572;
      W_f[14,8] := 0.14789321;
      W_f[14,9] := -0.08673888;
      W_f[14,10] := 0.41695347;
      W_f[14,11] := -0.40421456;
      W_f[14,12] := 0.20216350;
      W_f[14,13] := -0.08660001;
      W_f[14,14] := -0.07823719;
      W_f[14,15] := 0.32103771;
      W_f[14,16] := 0.02788324;
      W_f[14,17] := -0.09630302;
      W_f[14,18] := -0.54785252;
      W_f[14,19] := 0.17170331;
      W_f[14,20] := -0.17730309;
      W_f[14,21] := 0.29838467;
      W_f[14,22] := -0.17642282;
      W_f[14,23] := -0.04862199;
      W_f[14,24] := -1.37108374;
      W_f[14,25] := -0.24234977;
      W_f[14,26] := 0.08509517;
      W_f[14,27] := -0.30716902;
      W_f[14,28] := 0.77421099;
      W_f[14,29] := -0.42589924;
      W_f[14,30] := -0.18615769;
      W_f[14,31] := -0.12074227;
      W_f[14,32] := -0.08173326;
      W_f[14,33] := 0.03355461;
      W_f[14,34] := -0.12840785;
      W_f[14,35] := -0.04459246;
      W_f[14,36] := 0.08582738;
      W_f[14,37] := -0.03248604;
      W_f[14,38] := 0.00847942;
      W_f[14,39] := 0.16300382;
      W_f[15,0] := 0.03154271;
      W_f[15,1] := 0.05318842;
      W_f[15,2] := -0.10103899;
      W_f[15,3] := -0.02693522;
      W_f[15,4] := -0.06352412;
      W_f[15,5] := 0.09574427;
      W_f[15,6] := -0.03510033;
      W_f[15,7] := 0.01482865;
      W_f[15,8] := -0.02067289;
      W_f[15,9] := -0.04150250;
      W_f[15,10] := 0.01630465;
      W_f[15,11] := 0.06509072;
      W_f[15,12] := -0.17292246;
      W_f[15,13] := -0.11477651;
      W_f[15,14] := 0.23657221;
      W_f[15,15] := 0.09592439;
      W_f[15,16] := 0.07049410;
      W_f[15,17] := -0.04421110;
      W_f[15,18] := -0.17776524;
      W_f[15,19] := 0.06616033;
      W_f[15,20] := -0.05565001;
      W_f[15,21] := -0.05409446;
      W_f[15,22] := -0.05253718;
      W_f[15,23] := -0.06859960;
      W_f[15,24] := 0.02572974;
      W_f[15,25] := -0.02181539;
      W_f[15,26] := 0.00228037;
      W_f[15,27] := -0.05429837;
      W_f[15,28] := 0.06391250;
      W_f[15,29] := -0.05924486;
      W_f[15,30] := -0.09346493;
      W_f[15,31] := 0.02356213;
      W_f[15,32] := -0.07387451;
      W_f[15,33] := -0.15701193;
      W_f[15,34] := -0.50695050;
      W_f[15,35] := -0.11697226;
      W_f[15,36] := 0.03434648;
      W_f[15,37] := -0.08189469;
      W_f[15,38] := 0.22065248;
      W_f[15,39] := -0.17104173;
      W_f[16,0] := 0.17625535;
      W_f[16,1] := 0.11556054;
      W_f[16,2] := 0.07849861;
      W_f[16,3] := -0.34866714;
      W_f[16,4] := 0.03862548;
      W_f[16,5] := -0.22394647;
      W_f[16,6] := 0.11922321;
      W_f[16,7] := 0.13383812;
      W_f[16,8] := 0.12874119;
      W_f[16,9] := 0.11166555;
      W_f[16,10] := 0.03532283;
      W_f[16,11] := 0.12655254;
      W_f[16,12] := 0.15052819;
      W_f[16,13] := 0.01885046;
      W_f[16,14] := 0.57153022;
      W_f[16,15] := 0.22690293;
      W_f[16,16] := -0.22848204;
      W_f[16,17] := -0.40777546;
      W_f[16,18] := 0.18570280;
      W_f[16,19] := -0.50228417;
      W_f[16,20] := 0.07202365;
      W_f[16,21] := -0.02409742;
      W_f[16,22] := 0.03556022;
      W_f[16,23] := 0.25320294;
      W_f[16,24] := -0.85418850;
      W_f[16,25] := -0.75547177;
      W_f[16,26] := -0.01640177;
      W_f[16,27] := -0.22239800;
      W_f[16,28] := -0.06449725;
      W_f[16,29] := 0.12048583;
      W_f[16,30] := -0.09395292;
      W_f[16,31] := 0.14395721;
      W_f[16,32] := -0.37355945;
      W_f[16,33] := -0.22417888;
      W_f[16,34] := -1.13812256;
      W_f[16,35] := -0.22478914;
      W_f[16,36] := -0.00466719;
      W_f[16,37] := -0.22838083;
      W_f[16,38] := 0.13722458;
      W_f[16,39] := -0.27606511;
      W_f[17,0] := 0.09355596;
      W_f[17,1] := -0.03849373;
      W_f[17,2] := -0.22975640;
      W_f[17,3] := 0.05597479;
      W_f[17,4] := -0.12151184;
      W_f[17,5] := 0.09032618;
      W_f[17,6] := 0.05199543;
      W_f[17,7] := 0.09141852;
      W_f[17,8] := 0.09388466;
      W_f[17,9] := -0.00439828;
      W_f[17,10] := -0.17828138;
      W_f[17,11] := -0.35556960;
      W_f[17,12] := 0.37967008;
      W_f[17,13] := -0.08845654;
      W_f[17,14] := -0.07521001;
      W_f[17,15] := 0.00300852;
      W_f[17,16] := 0.08329321;
      W_f[17,17] := -0.09885437;
      W_f[17,18] := -0.00333220;
      W_f[17,19] := -0.31226391;
      W_f[17,20] := 0.22227764;
      W_f[17,21] := 0.37867606;
      W_f[17,22] := 0.17821352;
      W_f[17,23] := 0.00926425;
      W_f[17,24] := -0.15443780;
      W_f[17,25] := -0.39959320;
      W_f[17,26] := -0.10841592;
      W_f[17,27] := -0.36987418;
      W_f[17,28] := 0.09051982;
      W_f[17,29] := -0.11042830;
      W_f[17,30] := 0.06470256;
      W_f[17,31] := -0.06593291;
      W_f[17,32] := 0.33585012;
      W_f[17,33] := 0.47739133;
      W_f[17,34] := -1.25389719;
      W_f[17,35] := -0.16163990;
      W_f[17,36] := 0.07423314;
      W_f[17,37] := 0.00036682;
      W_f[17,38] := -0.11255764;
      W_f[17,39] := -0.06161462;
      W_f[18,0] := -0.04386483;
      W_f[18,1] := -0.10858835;
      W_f[18,2] := -0.28055254;
      W_f[18,3] := -0.04849620;
      W_f[18,4] := 0.12476673;
      W_f[18,5] := 0.10831297;
      W_f[18,6] := -0.08475895;
      W_f[18,7] := -0.18779263;
      W_f[18,8] := 0.01652613;
      W_f[18,9] := -0.02855963;
      W_f[18,10] := -0.06570389;
      W_f[18,11] := 0.06392785;
      W_f[18,12] := -0.08050973;
      W_f[18,13] := 0.05656723;
      W_f[18,14] := -0.02810039;
      W_f[18,15] := 0.15609136;
      W_f[18,16] := 0.14311801;
      W_f[18,17] := -0.09172881;
      W_f[18,18] := -0.18792967;
      W_f[18,19] := -0.40474713;
      W_f[18,20] := -0.30497348;
      W_f[18,21] := -0.42712539;
      W_f[18,22] := -0.07795502;
      W_f[18,23] := -0.17809948;
      W_f[18,24] := 0.20455103;
      W_f[18,25] := 0.01691615;
      W_f[18,26] := -0.35336512;
      W_f[18,27] := 0.11173917;
      W_f[18,28] := -0.10731182;
      W_f[18,29] := -0.06895053;
      W_f[18,30] := -0.08786953;
      W_f[18,31] := -0.19644345;
      W_f[18,32] := 0.07561095;
      W_f[18,33] := 0.13270301;
      W_f[18,34] := -0.00656677;
      W_f[18,35] := 0.11211497;
      W_f[18,36] := -0.13074799;
      W_f[18,37] := 0.07324994;
      W_f[18,38] := -0.00948287;
      W_f[18,39] := 0.08667010;
      W_f[19,0] := -0.05768050;
      W_f[19,1] := -0.00473207;
      W_f[19,2] := 0.09791042;
      W_f[19,3] := -0.02757404;
      W_f[19,4] := 0.16725993;
      W_f[19,5] := -0.00712524;
      W_f[19,6] := -0.02008255;
      W_f[19,7] := -0.05448977;
      W_f[19,8] := 0.00590254;
      W_f[19,9] := -0.10340165;
      W_f[19,10] := -0.02563939;
      W_f[19,11] := -0.07002047;
      W_f[19,12] := -0.00658451;
      W_f[19,13] := -0.06430968;
      W_f[19,14] := -0.24822524;
      W_f[19,15] := -0.27073550;
      W_f[19,16] := 0.10775120;
      W_f[19,17] := -0.19008251;
      W_f[19,18] := -0.14044385;
      W_f[19,19] := 0.91544735;
      W_f[19,20] := -0.07060743;
      W_f[19,21] := -0.01873856;
      W_f[19,22] := 0.08185165;
      W_f[19,23] := 0.06677809;
      W_f[19,24] := -0.63994950;
      W_f[19,25] := -0.76108485;
      W_f[19,26] := -0.12262011;
      W_f[19,27] := -0.13873395;
      W_f[19,28] := -0.12170569;
      W_f[19,29] := -0.13573299;
      W_f[19,30] := -0.02154119;
      W_f[19,31] := 0.13803685;
      W_f[19,32] := -0.25907481;
      W_f[19,33] := 0.00526916;
      W_f[19,34] := -1.01521635;
      W_f[19,35] := 0.00149761;
      W_f[19,36] := 0.01719889;
      W_f[19,37] := 0.06499543;
      W_f[19,38] := -0.31517512;
      W_f[19,39] := 0.79543614;
      W_f[20,0] := 0.16480501;
      W_f[20,1] := 0.08265622;
      W_f[20,2] := -0.23557226;
      W_f[20,3] := 0.55451566;
      W_f[20,4] := 0.01603219;
      W_f[20,5] := 0.04251210;
      W_f[20,6] := -0.11781015;
      W_f[20,7] := 0.01638467;
      W_f[20,8] := -0.83916026;
      W_f[20,9] := 0.24137184;
      W_f[20,10] := -0.33704534;
      W_f[20,11] := -0.12961838;
      W_f[20,12] := -0.06016191;
      W_f[20,13] := -0.07475966;
      W_f[20,14] := 0.06575783;
      W_f[20,15] := 0.22323456;
      W_f[20,16] := 0.13502784;
      W_f[20,17] := 0.00838923;
      W_f[20,18] := -0.10783752;
      W_f[20,19] := -0.13500038;
      W_f[20,20] := 0.08887729;
      W_f[20,21] := 0.10476577;
      W_f[20,22] := -0.28266746;
      W_f[20,23] := -0.20107298;
      W_f[20,24] := 1.60042787;
      W_f[20,25] := 1.42235684;
      W_f[20,26] := -0.10143545;
      W_f[20,27] := 0.21119232;
      W_f[20,28] := -0.12540008;
      W_f[20,29] := -0.08862077;
      W_f[20,30] := -0.16858271;
      W_f[20,31] := -0.37333480;
      W_f[20,32] := -0.28393903;
      W_f[20,33] := -0.27161008;
      W_f[20,34] := -0.08681910;
      W_f[20,35] := -0.17818987;
      W_f[20,36] := -0.03406080;
      W_f[20,37] := -0.08528435;
      W_f[20,38] := 0.03585081;
      W_f[20,39] := -0.18177070;
      W_f[21,0] := 0.04771005;
      W_f[21,1] := 0.08663736;
      W_f[21,2] := -0.02783780;
      W_f[21,3] := 0.07879353;
      W_f[21,4] := 0.27264851;
      W_f[21,5] := 0.07421625;
      W_f[21,6] := -0.12801333;
      W_f[21,7] := -0.08395027;
      W_f[21,8] := 0.04900100;
      W_f[21,9] := 0.20751640;
      W_f[21,10] := -0.32644811;
      W_f[21,11] := -0.06497382;
      W_f[21,12] := 0.09799027;
      W_f[21,13] := 0.00883581;
      W_f[21,14] := 0.00966343;
      W_f[21,15] := -0.14871061;
      W_f[21,16] := -0.00497553;
      W_f[21,17] := 0.11452187;
      W_f[21,18] := -0.20872478;
      W_f[21,19] := -0.10943013;
      W_f[21,20] := -0.18462080;
      W_f[21,21] := 0.05003940;
      W_f[21,22] := -0.13593008;
      W_f[21,23] := 0.03107853;
      W_f[21,24] := -0.04973240;
      W_f[21,25] := -0.15850165;
      W_f[21,26] := -0.04493616;
      W_f[21,27] := 0.06513418;
      W_f[21,28] := 0.02263425;
      W_f[21,29] := -0.14598361;
      W_f[21,30] := -0.20827983;
      W_f[21,31] := -0.22851680;
      W_f[21,32] := -0.16735223;
      W_f[21,33] := -0.15003826;
      W_f[21,34] := 0.11699387;
      W_f[21,35] := -0.04816795;
      W_f[21,36] := 0.06935357;
      W_f[21,37] := -0.10568924;
      W_f[21,38] := 0.03433881;
      W_f[21,39] := -0.05082455;
      W_f[22,0] := -0.21789505;
      W_f[22,1] := -0.00218185;
      W_f[22,2] := 0.13707796;
      W_f[22,3] := -0.05661480;
      W_f[22,4] := 0.04673120;
      W_f[22,5] := 0.07919453;
      W_f[22,6] := 0.00165318;
      W_f[22,7] := 0.24370010;
      W_f[22,8] := -0.49046701;
      W_f[22,9] := 0.18481795;
      W_f[22,10] := -0.09283270;
      W_f[22,11] := -0.08213542;
      W_f[22,12] := -0.11216073;
      W_f[22,13] := -0.12417459;
      W_f[22,14] := -0.03892196;
      W_f[22,15] := 0.00938558;
      W_f[22,16] := 0.04654559;
      W_f[22,17] := -0.01202954;
      W_f[22,18] := -0.08779050;
      W_f[22,19] := -0.04691886;
      W_f[22,20] := -0.04042359;
      W_f[22,21] := -0.10060240;
      W_f[22,22] := 0.30039361;
      W_f[22,23] := -0.14701439;
      W_f[22,24] := 0.92930299;
      W_f[22,25] := 0.95187950;
      W_f[22,26] := -0.14506029;
      W_f[22,27] := 0.09577515;
      W_f[22,28] := -0.03439396;
      W_f[22,29] := -0.13056463;
      W_f[22,30] := 0.23247777;
      W_f[22,31] := -0.01952458;
      W_f[22,32] := 0.29687238;
      W_f[22,33] := 0.05021480;
      W_f[22,34] := 0.61989981;
      W_f[22,35] := 0.12880597;
      W_f[22,36] := -0.00632370;
      W_f[22,37] := 0.26314035;
      W_f[22,38] := -0.13918042;
      W_f[22,39] := 0.48424563;
      W_f[23,0] := 0.18203287;
      W_f[23,1] := -0.00033453;
      W_f[23,2] := -0.12690647;
      W_f[23,3] := -0.20817837;
      W_f[23,4] := -0.03886449;
      W_f[23,5] := -0.07745034;
      W_f[23,6] := 0.09301028;
      W_f[23,7] := 0.29436016;
      W_f[23,8] := -0.00518724;
      W_f[23,9] := -0.06415172;
      W_f[23,10] := 0.09103597;
      W_f[23,11] := -0.11698931;
      W_f[23,12] := 0.04732081;
      W_f[23,13] := 0.04674791;
      W_f[23,14] := -0.02131645;
      W_f[23,15] := 0.04225742;
      W_f[23,16] := -0.17455494;
      W_f[23,17] := -0.03249518;
      W_f[23,18] := -0.30770859;
      W_f[23,19] := 0.33163178;
      W_f[23,20] := 0.14246757;
      W_f[23,21] := 0.14922017;
      W_f[23,22] := 0.15601201;
      W_f[23,23] := -0.00516094;
      W_f[23,24] := -1.45130980;
      W_f[23,25] := -0.36313021;
      W_f[23,26] := -0.07832589;
      W_f[23,27] := -0.16756825;
      W_f[23,28] := 0.07020092;
      W_f[23,29] := 0.15479565;
      W_f[23,30] := 0.18874301;
      W_f[23,31] := 0.02346863;
      W_f[23,32] := 0.01785002;
      W_f[23,33] := -0.12262850;
      W_f[23,34] := -0.04859183;
      W_f[23,35] := -0.14257406;
      W_f[23,36] := 0.00146115;
      W_f[23,37] := 0.09021772;
      W_f[23,38] := 0.14310881;
      W_f[23,39] := 0.10275228;
      W_f[24,0] := -0.05857223;
      W_f[24,1] := 0.15763901;
      W_f[24,2] := -0.13669187;
      W_f[24,3] := 0.13361017;
      W_f[24,4] := -0.01805840;
      W_f[24,5] := 0.08483858;
      W_f[24,6] := 0.06242542;
      W_f[24,7] := 0.09024160;
      W_f[24,8] := -0.02310267;
      W_f[24,9] := -0.21032517;
      W_f[24,10] := -0.05898380;
      W_f[24,11] := -0.07191398;
      W_f[24,12] := -0.17340270;
      W_f[24,13] := 0.05035622;
      W_f[24,14] := 0.11432620;
      W_f[24,15] := 0.09918343;
      W_f[24,16] := -0.09240849;
      W_f[24,17] := 0.06147276;
      W_f[24,18] := -0.15851578;
      W_f[24,19] := -0.19691418;
      W_f[24,20] := -0.06251538;
      W_f[24,21] := 0.09218568;
      W_f[24,22] := -0.03233892;
      W_f[24,23] := -0.13645050;
      W_f[24,24] := 1.50175047;
      W_f[24,25] := 1.34456754;
      W_f[24,26] := -0.00621613;
      W_f[24,27] := -0.01676605;
      W_f[24,28] := -0.02784773;
      W_f[24,29] := 0.62369519;
      W_f[24,30] := -0.12347586;
      W_f[24,31] := -0.03955586;
      W_f[24,32] := 0.14359131;
      W_f[24,33] := -0.02603620;
      W_f[24,34] := 1.24290085;
      W_f[24,35] := 0.02946699;
      W_f[24,36] := 0.23795766;
      W_f[24,37] := 0.14494100;
      W_f[24,38] := 0.14506596;
      W_f[24,39] := -0.03060411;
      W_f[25,0] := 0.04533798;
      W_f[25,1] := -0.07252404;
      W_f[25,2] := -0.04066183;
      W_f[25,3] := 0.19957697;
      W_f[25,4] := 0.03161494;
      W_f[25,5] := -0.03136744;
      W_f[25,6] := 0.02992978;
      W_f[25,7] := 0.01081558;
      W_f[25,8] := 0.18272607;
      W_f[25,9] := -0.01668218;
      W_f[25,10] := 0.01204226;
      W_f[25,11] := 0.07526124;
      W_f[25,12] := 0.03537060;
      W_f[25,13] := 0.10093886;
      W_f[25,14] := -0.12508741;
      W_f[25,15] := -0.04653997;
      W_f[25,16] := 0.00332855;
      W_f[25,17] := 0.03725290;
      W_f[25,18] := -0.09655500;
      W_f[25,19] := -0.30870706;
      W_f[25,20] := -0.10335279;
      W_f[25,21] := -0.19976620;
      W_f[25,22] := -0.03147923;
      W_f[25,23] := -0.14786926;
      W_f[25,24] := -0.27878088;
      W_f[25,25] := -0.34400648;
      W_f[25,26] := -0.21661498;
      W_f[25,27] := 0.29630589;
      W_f[25,28] := 0.03365128;
      W_f[25,29] := 0.22238778;
      W_f[25,30] := 0.10650972;
      W_f[25,31] := -0.10210063;
      W_f[25,32] := 0.14446351;
      W_f[25,33] := 0.02928571;
      W_f[25,34] := -0.11391223;
      W_f[25,35] := 0.11920016;
      W_f[25,36] := -0.11559187;
      W_f[25,37] := 0.19095075;
      W_f[25,38] := -0.04105619;
      W_f[25,39] := 0.23975134;
      W_f[26,0] := 0.00493505;
      W_f[26,1] := 0.07623698;
      W_f[26,2] := -0.01626105;
      W_f[26,3] := 0.08502831;
      W_f[26,4] := 0.11989306;
      W_f[26,5] := 0.05587002;
      W_f[26,6] := -0.23084743;
      W_f[26,7] := -0.17441489;
      W_f[26,8] := 0.00085686;
      W_f[26,9] := -0.05871731;
      W_f[26,10] := 0.07582050;
      W_f[26,11] := -0.19967213;
      W_f[26,12] := -0.31389868;
      W_f[26,13] := 0.13419744;
      W_f[26,14] := 0.02738570;
      W_f[26,15] := -0.04184799;
      W_f[26,16] := 0.02028807;
      W_f[26,17] := 0.00563849;
      W_f[26,18] := -0.12281100;
      W_f[26,19] := 0.00383526;
      W_f[26,20] := -0.06410136;
      W_f[26,21] := -0.06429290;
      W_f[26,22] := -0.08350200;
      W_f[26,23] := -0.10770558;
      W_f[26,24] := 0.45600012;
      W_f[26,25] := 0.27628049;
      W_f[26,26] := -0.01219090;
      W_f[26,27] := 0.09856915;
      W_f[26,28] := 0.08391341;
      W_f[26,29] := -0.15169400;
      W_f[26,30] := -0.05663548;
      W_f[26,31] := 0.01523839;
      W_f[26,32] := -0.00722656;
      W_f[26,33] := 0.00556829;
      W_f[26,34] := -0.39934179;
      W_f[26,35] := -0.04286478;
      W_f[26,36] := -0.01076956;
      W_f[26,37] := -0.02061651;
      W_f[26,38] := 0.13584487;
      W_f[26,39] := 0.01977600;
      W_f[27,0] := -0.10016902;
      W_f[27,1] := 0.07916581;
      W_f[27,2] := 0.15547076;
      W_f[27,3] := 0.70207226;
      W_f[27,4] := -0.00100257;
      W_f[27,5] := 0.16907251;
      W_f[27,6] := 0.09067014;
      W_f[27,7] := -0.48238862;
      W_f[27,8] := -0.32165852;
      W_f[27,9] := -0.15741454;
      W_f[27,10] := -0.14824116;
      W_f[27,11] := -0.00698989;
      W_f[27,12] := -0.11109005;
      W_f[27,13] := -0.24554738;
      W_f[27,14] := 0.04736808;
      W_f[27,15] := 0.14338875;
      W_f[27,16] := -0.10880961;
      W_f[27,17] := 0.09295370;
      W_f[27,18] := -0.13496843;
      W_f[27,19] := -0.17531624;
      W_f[27,20] := -0.01208391;
      W_f[27,21] := -0.21940263;
      W_f[27,22] := -0.14602076;
      W_f[27,23] := -0.04240515;
      W_f[27,24] := 1.45130336;
      W_f[27,25] := 1.26312649;
      W_f[27,26] := -0.06854503;
      W_f[27,27] := 0.11704011;
      W_f[27,28] := 0.09159904;
      W_f[27,29] := -0.04047090;
      W_f[27,30] := -0.10142513;
      W_f[27,31] := -0.03332018;
      W_f[27,32] := -0.03741011;
      W_f[27,33] := -0.02919200;
      W_f[27,34] := -0.21617067;
      W_f[27,35] := -0.15822560;
      W_f[27,36] := 0.15107271;
      W_f[27,37] := -0.00820841;
      W_f[27,38] := 0.05202204;
      W_f[27,39] := -0.08140420;
      W_f[28,0] := 0.21725248;
      W_f[28,1] := 0.11601064;
      W_f[28,2] := -0.50731003;
      W_f[28,3] := 0.34125856;
      W_f[28,4] := 0.01358903;
      W_f[28,5] := 0.07589430;
      W_f[28,6] := 0.14723879;
      W_f[28,7] := 0.04250083;
      W_f[28,8] := -0.74850899;
      W_f[28,9] := 0.35015193;
      W_f[28,10] := 0.02476582;
      W_f[28,11] := -0.08709566;
      W_f[28,12] := -0.14858241;
      W_f[28,13] := 0.10917792;
      W_f[28,14] := -0.01036290;
      W_f[28,15] := -0.00310236;
      W_f[28,16] := -0.11779232;
      W_f[28,17] := -0.09907542;
      W_f[28,18] := 0.04596486;
      W_f[28,19] := 0.02090520;
      W_f[28,20] := 0.04032231;
      W_f[28,21] := -0.02343630;
      W_f[28,22] := 0.31838682;
      W_f[28,23] := -0.18608692;
      W_f[28,24] := 1.11693740;
      W_f[28,25] := 1.13061082;
      W_f[28,26] := -0.01059407;
      W_f[28,27] := 0.04070573;
      W_f[28,28] := 0.23042743;
      W_f[28,29] := 0.39798027;
      W_f[28,30] := 0.31331325;
      W_f[28,31] := 0.01896788;
      W_f[28,32] := 0.05937084;
      W_f[28,33] := 0.32739767;
      W_f[28,34] := 0.11175870;
      W_f[28,35] := 0.38728848;
      W_f[28,36] := 0.07428543;
      W_f[28,37] := 0.28699094;
      W_f[28,38] := 0.02707092;
      W_f[28,39] := 0.09776948;
      W_f[29,0] := -0.05480788;
      W_f[29,1] := -0.06971346;
      W_f[29,2] := 0.15541564;
      W_f[29,3] := -0.02117513;
      W_f[29,4] := -0.02765184;
      W_f[29,5] := 0.48948473;
      W_f[29,6] := 0.23739967;
      W_f[29,7] := 0.39359435;
      W_f[29,8] := 0.12403622;
      W_f[29,9] := -0.23649004;
      W_f[29,10] := 0.21631436;
      W_f[29,11] := -0.22992733;
      W_f[29,12] := -0.11843852;
      W_f[29,13] := 0.12832482;
      W_f[29,14] := 0.15944116;
      W_f[29,15] := 0.16688094;
      W_f[29,16] := -0.03219134;
      W_f[29,17] := 0.07033925;
      W_f[29,18] := 0.15342207;
      W_f[29,19] := -0.08973140;
      W_f[29,20] := 0.01753044;
      W_f[29,21] := -0.21804836;
      W_f[29,22] := 0.10274304;
      W_f[29,23] := -0.07748783;
      W_f[29,24] := 0.14996310;
      W_f[29,25] := 0.05747431;
      W_f[29,26] := -0.05352241;
      W_f[29,27] := 0.20547068;
      W_f[29,28] := 0.21826106;
      W_f[29,29] := -0.49819168;
      W_f[29,30] := -0.07471830;
      W_f[29,31] := -0.12761955;
      W_f[29,32] := -0.08077794;
      W_f[29,33] := 0.16914612;
      W_f[29,34] := -0.02049359;
      W_f[29,35] := -0.25413868;
      W_f[29,36] := -0.03029504;
      W_f[29,37] := -0.04286458;
      W_f[29,38] := -0.00078733;
      W_f[29,39] := 0.06210590;
      W_f[30,0] := 0.04379491;
      W_f[30,1] := -0.06586411;
      W_f[30,2] := -0.13123371;
      W_f[30,3] := -0.37808374;
      W_f[30,4] := 0.10017996;
      W_f[30,5] := -0.03991124;
      W_f[30,6] := 0.04357130;
      W_f[30,7] := -0.18068686;
      W_f[30,8] := -0.00580577;
      W_f[30,9] := 0.36891636;
      W_f[30,10] := 0.01027874;
      W_f[30,11] := 0.50609785;
      W_f[30,12] := 0.01925549;
      W_f[30,13] := -0.06952953;
      W_f[30,14] := 0.03735949;
      W_f[30,15] := -0.85169780;
      W_f[30,16] := -0.14351282;
      W_f[30,17] := 0.09829179;
      W_f[30,18] := 0.13755107;
      W_f[30,19] := 0.14171647;
      W_f[30,20] := 0.15322028;
      W_f[30,21] := -0.01534852;
      W_f[30,22] := -0.07220063;
      W_f[30,23] := -0.00489338;
      W_f[30,24] := -0.08854904;
      W_f[30,25] := 0.11646047;
      W_f[30,26] := -0.04590597;
      W_f[30,27] := -0.12970480;
      W_f[30,28] := 0.03094332;
      W_f[30,29] := 0.33986101;
      W_f[30,30] := -0.11265934;
      W_f[30,31] := -0.00355576;
      W_f[30,32] := -0.07702769;
      W_f[30,33] := -0.03350009;
      W_f[30,34] := 0.04180816;
      W_f[30,35] := -0.01911464;
      W_f[30,36] := 0.01183037;
      W_f[30,37] := 0.22970138;
      W_f[30,38] := 0.01091551;
      W_f[30,39] := -0.10615819;
      W_f[31,0] := -0.12645298;
      W_f[31,1] := -0.03490535;
      W_f[31,2] := -0.04712384;
      W_f[31,3] := -0.22141387;
      W_f[31,4] := -0.06836447;
      W_f[31,5] := 0.15984270;
      W_f[31,6] := 0.04255423;
      W_f[31,7] := -0.03223060;
      W_f[31,8] := 0.02700607;
      W_f[31,9] := -0.09661999;
      W_f[31,10] := 0.15196519;
      W_f[31,11] := -0.03100767;
      W_f[31,12] := 0.06127577;
      W_f[31,13] := 0.00739274;
      W_f[31,14] := 0.00656646;
      W_f[31,15] := 0.16660002;
      W_f[31,16] := 0.32314840;
      W_f[31,17] := 0.00930041;
      W_f[31,18] := 0.02132557;
      W_f[31,19] := 0.00431878;
      W_f[31,20] := 0.06450959;
      W_f[31,21] := 0.08898797;
      W_f[31,22] := 0.14660980;
      W_f[31,23] := 0.00585541;
      W_f[31,24] := 0.55362934;
      W_f[31,25] := 0.56018978;
      W_f[31,26] := -0.09814498;
      W_f[31,27] := -0.02094743;
      W_f[31,28] := 0.07426088;
      W_f[31,29] := 0.38328037;
      W_f[31,30] := 0.32430744;
      W_f[31,31] := -0.26375374;
      W_f[31,32] := 0.26633716;
      W_f[31,33] := 0.01791180;
      W_f[31,34] := -0.01126823;
      W_f[31,35] := 0.15723105;
      W_f[31,36] := 0.04929269;
      W_f[31,37] := 0.41218692;
      W_f[31,38] := 0.01116225;
      W_f[31,39] := 0.14782998;
      W_g[0,0] := -0.29731244;
      W_g[0,1] := 0.30804923;
      W_g[0,2] := -0.07333095;
      W_g[0,3] := 0.21897507;
      W_g[0,4] := -0.21115625;
      W_g[0,5] := 0.04973322;
      W_g[0,6] := -0.18843463;
      W_g[0,7] := 0.13841841;
      W_g[0,8] := 0.18074706;
      W_g[0,9] := 0.13372360;
      W_g[0,10] := -0.22122957;
      W_g[0,11] := -0.34522530;
      W_g[0,12] := 0.07657024;
      W_g[0,13] := 0.11239351;
      W_g[0,14] := 0.00508291;
      W_g[0,15] := 0.00489822;
      W_g[0,16] := -0.04131620;
      W_g[0,17] := -0.07313628;
      W_g[0,18] := 0.03842196;
      W_g[0,19] := 0.31408229;
      W_g[0,20] := 0.14011617;
      W_g[0,21] := -0.27653301;
      W_g[0,22] := -0.09168060;
      W_g[0,23] := 0.22705604;
      W_g[0,24] := 0.51337552;
      W_g[0,25] := 0.55914593;
      W_g[0,26] := 0.33094329;
      W_g[0,27] := 0.20361137;
      W_g[0,28] := -0.03624717;
      W_g[0,29] := 0.08691628;
      W_g[0,30] := -0.08794427;
      W_g[0,31] := -0.15352608;
      W_g[0,32] := 0.05986316;
      W_g[0,33] := 0.05109673;
      W_g[0,34] := 0.67403698;
      W_g[0,35] := 0.15075700;
      W_g[0,36] := 0.00786592;
      W_g[0,37] := 0.17828523;
      W_g[0,38] := 0.15761673;
      W_g[0,39] := 0.00874934;
      W_g[1,0] := 0.32671660;
      W_g[1,1] := 0.01836558;
      W_g[1,2] := 0.25563437;
      W_g[1,3] := 0.14020202;
      W_g[1,4] := 0.13369501;
      W_g[1,5] := -0.06653731;
      W_g[1,6] := 0.07586989;
      W_g[1,7] := 0.19387591;
      W_g[1,8] := 0.26986131;
      W_g[1,9] := 0.27328917;
      W_g[1,10] := 0.20197332;
      W_g[1,11] := 0.05846954;
      W_g[1,12] := 0.10516258;
      W_g[1,13] := -0.10580415;
      W_g[1,14] := -0.00597053;
      W_g[1,15] := -0.00393197;
      W_g[1,16] := -0.00673947;
      W_g[1,17] := -0.03512664;
      W_g[1,18] := -0.04886592;
      W_g[1,19] := -0.00479484;
      W_g[1,20] := 0.15406653;
      W_g[1,21] := 0.04567941;
      W_g[1,22] := -0.01350505;
      W_g[1,23] := 0.02950142;
      W_g[1,24] := 0.01168221;
      W_g[1,25] := 0.35458666;
      W_g[1,26] := 0.03195773;
      W_g[1,27] := 0.04014106;
      W_g[1,28] := 0.04925289;
      W_g[1,29] := -0.04943694;
      W_g[1,30] := -0.02163855;
      W_g[1,31] := -0.02884842;
      W_g[1,32] := -0.02839119;
      W_g[1,33] := -0.03380399;
      W_g[1,34] := 0.19551215;
      W_g[1,35] := -0.02271999;
      W_g[1,36] := -0.01233778;
      W_g[1,37] := 0.01909558;
      W_g[1,38] := -0.02520212;
      W_g[1,39] := -0.03295163;
      W_g[2,0] := -0.15581730;
      W_g[2,1] := 0.01425133;
      W_g[2,2] := 0.13872904;
      W_g[2,3] := -0.13885449;
      W_g[2,4] := -0.29651093;
      W_g[2,5] := 0.06956124;
      W_g[2,6] := 0.23148759;
      W_g[2,7] := 0.10803487;
      W_g[2,8] := -0.02653480;
      W_g[2,9] := 0.17615019;
      W_g[2,10] := -0.15386169;
      W_g[2,11] := -0.12791342;
      W_g[2,12] := -0.16833690;
      W_g[2,13] := -0.02681257;
      W_g[2,14] := -0.04338213;
      W_g[2,15] := -0.00641101;
      W_g[2,16] := -0.01647951;
      W_g[2,17] := -0.10473385;
      W_g[2,18] := 0.02287934;
      W_g[2,19] := 0.01147376;
      W_g[2,20] := -0.07240344;
      W_g[2,21] := 0.18736833;
      W_g[2,22] := -0.09113216;
      W_g[2,23] := -0.05816693;
      W_g[2,24] := -0.09419736;
      W_g[2,25] := -0.23981659;
      W_g[2,26] := 0.03237080;
      W_g[2,27] := 0.58103901;
      W_g[2,28] := 0.68347645;
      W_g[2,29] := -0.06846042;
      W_g[2,30] := -0.08991379;
      W_g[2,31] := -0.06568053;
      W_g[2,32] := -0.00146176;
      W_g[2,33] := -0.05521696;
      W_g[2,34] := -0.27966231;
      W_g[2,35] := 0.07491860;
      W_g[2,36] := -0.16886964;
      W_g[2,37] := 0.07337529;
      W_g[2,38] := 0.02869449;
      W_g[2,39] := -0.05087301;
      W_g[3,0] := 0.21261550;
      W_g[3,1] := 0.07068379;
      W_g[3,2] := 0.23964408;
      W_g[3,3] := 0.25374594;
      W_g[3,4] := -0.07897907;
      W_g[3,5] := 0.53360569;
      W_g[3,6] := -0.50441998;
      W_g[3,7] := -0.43295726;
      W_g[3,8] := 0.45935890;
      W_g[3,9] := -0.16401440;
      W_g[3,10] := -0.56816226;
      W_g[3,11] := 0.84965134;
      W_g[3,12] := 0.37320843;
      W_g[3,13] := 0.37158751;
      W_g[3,14] := 0.59009206;
      W_g[3,15] := -0.01866211;
      W_g[3,16] := -0.12090266;
      W_g[3,17] := -0.23170036;
      W_g[3,18] := -0.20994744;
      W_g[3,19] := -0.75220180;
      W_g[3,20] := 0.19406919;
      W_g[3,21] := -0.19833040;
      W_g[3,22] := -0.13843380;
      W_g[3,23] := -0.08076543;
      W_g[3,24] := -0.02181598;
      W_g[3,25] := 0.06219065;
      W_g[3,26] := -0.09015898;
      W_g[3,27] := 0.17478789;
      W_g[3,28] := 0.03573907;
      W_g[3,29] := 0.03600015;
      W_g[3,30] := -0.15354984;
      W_g[3,31] := 0.19793989;
      W_g[3,32] := 0.02940232;
      W_g[3,33] := -0.01058361;
      W_g[3,34] := 0.20539114;
      W_g[3,35] := 0.00076983;
      W_g[3,36] := -0.04329271;
      W_g[3,37] := 0.19885710;
      W_g[3,38] := -0.08021279;
      W_g[3,39] := 0.97782809;
      W_g[4,0] := -0.16564122;
      W_g[4,1] := -0.11781788;
      W_g[4,2] := 0.16660716;
      W_g[4,3] := -0.08943526;
      W_g[4,4] := 0.12463316;
      W_g[4,5] := 0.02390479;
      W_g[4,6] := -0.05541207;
      W_g[4,7] := -0.14321095;
      W_g[4,8] := -0.05963109;
      W_g[4,9] := -0.13049991;
      W_g[4,10] := 0.28670028;
      W_g[4,11] := -0.03267299;
      W_g[4,12] := -0.08092957;
      W_g[4,13] := -0.42708814;
      W_g[4,14] := -0.00459089;
      W_g[4,15] := 0.05856811;
      W_g[4,16] := 0.03812011;
      W_g[4,17] := -0.00688081;
      W_g[4,18] := 0.03390410;
      W_g[4,19] := 0.01956543;
      W_g[4,20] := 0.20069234;
      W_g[4,21] := -0.01636098;
      W_g[4,22] := 0.01006647;
      W_g[4,23] := 0.84444892;
      W_g[4,24] := 0.00210755;
      W_g[4,25] := -0.06413154;
      W_g[4,26] := -0.45401627;
      W_g[4,27] := 0.25349951;
      W_g[4,28] := -0.09389957;
      W_g[4,29] := 0.07596151;
      W_g[4,30] := 0.13383749;
      W_g[4,31] := 0.33215305;
      W_g[4,32] := 0.20357370;
      W_g[4,33] := 0.12820803;
      W_g[4,34] := 0.00518544;
      W_g[4,35] := 0.08931676;
      W_g[4,36] := -0.01421158;
      W_g[4,37] := 0.20269936;
      W_g[4,38] := 0.08788820;
      W_g[4,39] := -0.01560517;
      W_g[5,0] := -0.08699985;
      W_g[5,1] := 0.66933864;
      W_g[5,2] := -0.00633939;
      W_g[5,3] := -0.17376915;
      W_g[5,4] := 0.02668794;
      W_g[5,5] := -0.08880353;
      W_g[5,6] := -0.11177815;
      W_g[5,7] := 0.26541734;
      W_g[5,8] := -0.09973598;
      W_g[5,9] := 0.29554251;
      W_g[5,10] := -0.37329444;
      W_g[5,11] := 0.09036310;
      W_g[5,12] := -0.29482436;
      W_g[5,13] := -0.35888001;
      W_g[5,14] := -0.01915385;
      W_g[5,15] := 0.04767168;
      W_g[5,16] := 0.03428055;
      W_g[5,17] := 0.03784378;
      W_g[5,18] := 0.04297538;
      W_g[5,19] := -0.24454381;
      W_g[5,20] := -0.34855694;
      W_g[5,21] := -0.15681590;
      W_g[5,22] := 0.04547088;
      W_g[5,23] := -0.15585004;
      W_g[5,24] := 0.01251255;
      W_g[5,25] := 0.15953992;
      W_g[5,26] := -0.18765861;
      W_g[5,27] := -0.01743420;
      W_g[5,28] := -0.23351699;
      W_g[5,29] := 0.02074986;
      W_g[5,30] := 0.02202098;
      W_g[5,31] := 0.24873479;
      W_g[5,32] := 0.06216014;
      W_g[5,33] := 0.06517217;
      W_g[5,34] := 0.02405161;
      W_g[5,35] := 0.04143449;
      W_g[5,36] := 0.08146483;
      W_g[5,37] := 0.16652697;
      W_g[5,38] := 0.01448802;
      W_g[5,39] := 0.08552948;
      W_g[6,0] := -0.14679314;
      W_g[6,1] := 0.04948491;
      W_g[6,2] := 0.02849484;
      W_g[6,3] := -0.08913121;
      W_g[6,4] := 0.01332707;
      W_g[6,5] := 0.02870432;
      W_g[6,6] := -0.13538505;
      W_g[6,7] := 0.10151362;
      W_g[6,8] := 0.07108080;
      W_g[6,9] := 0.15849109;
      W_g[6,10] := -0.22181113;
      W_g[6,11] := -0.03935358;
      W_g[6,12] := 0.04531641;
      W_g[6,13] := 0.10437059;
      W_g[6,14] := 0.00934802;
      W_g[6,15] := -0.00473133;
      W_g[6,16] := 0.19776262;
      W_g[6,17] := 0.06397073;
      W_g[6,18] := -0.08264492;
      W_g[6,19] := -0.00858563;
      W_g[6,20] := 0.59372175;
      W_g[6,21] := -0.02809042;
      W_g[6,22] := 0.01213905;
      W_g[6,23] := -0.10024478;
      W_g[6,24] := -0.24557531;
      W_g[6,25] := -0.05298537;
      W_g[6,26] := -0.16861317;
      W_g[6,27] := 0.08932645;
      W_g[6,28] := 0.15916736;
      W_g[6,29] := -0.06639078;
      W_g[6,30] := 0.01585412;
      W_g[6,31] := 0.54062325;
      W_g[6,32] := -0.15765822;
      W_g[6,33] := -0.16314203;
      W_g[6,34] := -0.18088351;
      W_g[6,35] := -0.25276086;
      W_g[6,36] := -0.02972133;
      W_g[6,37] := -0.22347295;
      W_g[6,38] := 0.12736996;
      W_g[6,39] := 0.02743512;
      W_g[7,0] := -0.16503690;
      W_g[7,1] := 0.03972364;
      W_g[7,2] := -0.00654130;
      W_g[7,3] := 0.47248334;
      W_g[7,4] := 0.22141388;
      W_g[7,5] := -0.02702056;
      W_g[7,6] := -0.08594248;
      W_g[7,7] := -0.10240269;
      W_g[7,8] := 0.08587579;
      W_g[7,9] := -0.29143050;
      W_g[7,10] := -0.04244880;
      W_g[7,11] := 0.07958402;
      W_g[7,12] := 0.05996885;
      W_g[7,13] := 0.04256921;
      W_g[7,14] := 0.14755034;
      W_g[7,15] := -0.13249832;
      W_g[7,16] := -0.02742708;
      W_g[7,17] := 0.07044590;
      W_g[7,18] := -0.01704550;
      W_g[7,19] := 0.11561061;
      W_g[7,20] := -0.04334126;
      W_g[7,21] := 0.30209017;
      W_g[7,22] := 0.12059546;
      W_g[7,23] := -0.01143128;
      W_g[7,24] := 0.43696722;
      W_g[7,25] := 0.27256724;
      W_g[7,26] := -0.01071244;
      W_g[7,27] := -0.05641021;
      W_g[7,28] := -0.11184577;
      W_g[7,29] := -0.12506962;
      W_g[7,30] := 0.11383872;
      W_g[7,31] := -0.12637268;
      W_g[7,32] := 0.01232483;
      W_g[7,33] := -0.05794921;
      W_g[7,34] := 0.14192834;
      W_g[7,35] := 0.04089052;
      W_g[7,36] := -0.26191169;
      W_g[7,37] := 0.00023886;
      W_g[7,38] := 0.00715496;
      W_g[7,39] := 0.08836767;
      W_g[8,0] := 0.12069551;
      W_g[8,1] := -0.05102030;
      W_g[8,2] := -0.08442411;
      W_g[8,3] := -0.16018370;
      W_g[8,4] := -0.03896859;
      W_g[8,5] := 0.00796033;
      W_g[8,6] := 0.03281215;
      W_g[8,7] := 0.04158888;
      W_g[8,8] := -0.06430040;
      W_g[8,9] := 0.13734795;
      W_g[8,10] := 0.03013904;
      W_g[8,11] := -0.19144072;
      W_g[8,12] := 0.18297645;
      W_g[8,13] := -0.02042261;
      W_g[8,14] := 0.47640336;
      W_g[8,15] := -0.07802652;
      W_g[8,16] := 0.03107872;
      W_g[8,17] := -0.09448601;
      W_g[8,18] := 0.02560257;
      W_g[8,19] := 0.24542020;
      W_g[8,20] := 0.01119845;
      W_g[8,21] := -0.30462247;
      W_g[8,22] := -0.04350797;
      W_g[8,23] := -0.16951585;
      W_g[8,24] := 0.12095571;
      W_g[8,25] := 0.08566401;
      W_g[8,26] := -0.13064992;
      W_g[8,27] := 0.16942461;
      W_g[8,28] := -0.00051321;
      W_g[8,29] := -0.16719460;
      W_g[8,30] := -0.03225356;
      W_g[8,31] := 0.16128831;
      W_g[8,32] := 0.05924257;
      W_g[8,33] := 0.06252825;
      W_g[8,34] := 0.04885080;
      W_g[8,35] := 0.06716868;
      W_g[8,36] := -0.02168992;
      W_g[8,37] := 0.08623782;
      W_g[8,38] := -0.06822046;
      W_g[8,39] := -0.03733813;
      W_g[9,0] := 0.81871593;
      W_g[9,1] := 0.02526643;
      W_g[9,2] := -0.76041377;
      W_g[9,3] := 0.51836115;
      W_g[9,4] := -0.21780470;
      W_g[9,5] := 0.02361593;
      W_g[9,6] := -0.55600011;
      W_g[9,7] := 0.06145347;
      W_g[9,8] := 0.04358738;
      W_g[9,9] := -0.21609305;
      W_g[9,10] := -0.10566008;
      W_g[9,11] := -0.00301302;
      W_g[9,12] := 0.35560456;
      W_g[9,13] := -0.22366437;
      W_g[9,14] := -0.00890417;
      W_g[9,15] := 0.31469098;
      W_g[9,16] := 0.14210188;
      W_g[9,17] := 0.32488760;
      W_g[9,18] := -0.10977074;
      W_g[9,19] := -0.22636354;
      W_g[9,20] := -0.32791817;
      W_g[9,21] := -0.57256800;
      W_g[9,22] := -0.28585047;
      W_g[9,23] := 0.20341209;
      W_g[9,24] := -0.76711357;
      W_g[9,25] := -0.89817464;
      W_g[9,26] := -0.32050338;
      W_g[9,27] := 0.39106333;
      W_g[9,28] := 0.43121040;
      W_g[9,29] := 0.14572853;
      W_g[9,30] := -0.16380118;
      W_g[9,31] := -0.30435774;
      W_g[9,32] := -0.06825320;
      W_g[9,33] := -0.15947679;
      W_g[9,34] := -0.12722060;
      W_g[9,35] := 0.27286705;
      W_g[9,36] := -0.17627911;
      W_g[9,37] := 0.20060076;
      W_g[9,38] := -0.23259346;
      W_g[9,39] := -0.20107704;
      W_g[10,0] := -0.03653082;
      W_g[10,1] := -0.00459500;
      W_g[10,2] := 0.04608782;
      W_g[10,3] := -0.08378540;
      W_g[10,4] := -0.00994155;
      W_g[10,5] := 0.10961147;
      W_g[10,6] := 0.15406886;
      W_g[10,7] := -0.11930396;
      W_g[10,8] := -0.00437860;
      W_g[10,9] := 0.05714689;
      W_g[10,10] := -0.00173966;
      W_g[10,11] := -0.57551277;
      W_g[10,12] := 0.42625594;
      W_g[10,13] := -0.40591905;
      W_g[10,14] := -0.19576681;
      W_g[10,15] := 0.08438285;
      W_g[10,16] := -0.01722066;
      W_g[10,17] := 0.04172579;
      W_g[10,18] := -0.06110490;
      W_g[10,19] := 0.08427376;
      W_g[10,20] := -0.10799333;
      W_g[10,21] := -0.00058548;
      W_g[10,22] := 0.06713647;
      W_g[10,23] := -0.09210554;
      W_g[10,24] := -0.09937313;
      W_g[10,25] := -0.07247933;
      W_g[10,26] := 0.20139590;
      W_g[10,27] := -0.03532998;
      W_g[10,28] := -0.08083174;
      W_g[10,29] := 0.21411720;
      W_g[10,30] := 0.01127313;
      W_g[10,31] := -0.06344012;
      W_g[10,32] := 0.02854561;
      W_g[10,33] := 0.02152516;
      W_g[10,34] := 0.00244472;
      W_g[10,35] := -0.11918493;
      W_g[10,36] := -0.00852005;
      W_g[10,37] := 0.05143885;
      W_g[10,38] := -0.03254176;
      W_g[10,39] := 0.62638599;
      W_g[11,0] := 0.13177699;
      W_g[11,1] := -0.06769224;
      W_g[11,2] := 0.10452202;
      W_g[11,3] := 0.05449197;
      W_g[11,4] := 0.01810149;
      W_g[11,5] := 0.03084538;
      W_g[11,6] := -0.02990450;
      W_g[11,7] := -0.02282630;
      W_g[11,8] := -0.17183347;
      W_g[11,9] := -0.11026753;
      W_g[11,10] := 0.08694904;
      W_g[11,11] := -0.08632144;
      W_g[11,12] := 0.15890475;
      W_g[11,13] := 0.15897611;
      W_g[11,14] := -0.06856292;
      W_g[11,15] := 0.12105770;
      W_g[11,16] := -0.03902842;
      W_g[11,17] := 0.15743148;
      W_g[11,18] := -0.05494931;
      W_g[11,19] := -0.31661710;
      W_g[11,20] := 0.00237431;
      W_g[11,21] := -0.29374212;
      W_g[11,22] := -0.00387868;
      W_g[11,23] := -0.15384512;
      W_g[11,24] := 0.26705560;
      W_g[11,25] := 0.28627306;
      W_g[11,26] := 0.16300470;
      W_g[11,27] := 0.36486325;
      W_g[11,28] := -0.10527802;
      W_g[11,29] := -0.06614047;
      W_g[11,30] := 0.00622322;
      W_g[11,31] := 0.31526664;
      W_g[11,32] := 0.06752055;
      W_g[11,33] := 0.00520946;
      W_g[11,34] := 0.01956053;
      W_g[11,35] := 0.03621605;
      W_g[11,36] := -0.11561473;
      W_g[11,37] := 0.09378653;
      W_g[11,38] := 0.06442897;
      W_g[11,39] := -0.06822205;
      W_g[12,0] := -0.34109655;
      W_g[12,1] := -0.06000578;
      W_g[12,2] := -0.09373351;
      W_g[12,3] := 0.08326271;
      W_g[12,4] := 0.00906463;
      W_g[12,5] := 0.07884520;
      W_g[12,6] := 0.05942823;
      W_g[12,7] := 0.28550220;
      W_g[12,8] := -0.36121264;
      W_g[12,9] := 0.12771368;
      W_g[12,10] := 0.03765302;
      W_g[12,11] := 0.13665034;
      W_g[12,12] := 0.35631377;
      W_g[12,13] := -0.21096121;
      W_g[12,14] := -0.02360137;
      W_g[12,15] := 0.15230067;
      W_g[12,16] := -0.00824362;
      W_g[12,17] := -0.09702953;
      W_g[12,18] := -0.26124185;
      W_g[12,19] := -0.19844258;
      W_g[12,20] := 0.10597581;
      W_g[12,21] := -0.12326175;
      W_g[12,22] := -0.01443423;
      W_g[12,23] := -0.02930082;
      W_g[12,24] := 0.18288726;
      W_g[12,25] := 0.19803882;
      W_g[12,26] := 0.04977860;
      W_g[12,27] := 0.04707592;
      W_g[12,28] := 0.04168066;
      W_g[12,29] := -0.11191346;
      W_g[12,30] := -0.00637640;
      W_g[12,31] := -0.05627256;
      W_g[12,32] := 0.04867624;
      W_g[12,33] := 0.02836183;
      W_g[12,34] := 0.29845282;
      W_g[12,35] := 0.07853222;
      W_g[12,36] := 0.01144999;
      W_g[12,37] := 0.03406933;
      W_g[12,38] := -0.05539230;
      W_g[12,39] := 0.04716556;
      W_g[13,0] := -0.06528508;
      W_g[13,1] := 0.04750456;
      W_g[13,2] := 0.00729868;
      W_g[13,3] := 0.19038309;
      W_g[13,4] := -0.26934335;
      W_g[13,5] := 0.07256790;
      W_g[13,6] := -0.04099108;
      W_g[13,7] := -0.02624341;
      W_g[13,8] := -0.05020488;
      W_g[13,9] := -0.10872720;
      W_g[13,10] := -0.06591415;
      W_g[13,11] := -0.14674501;
      W_g[13,12] := 0.20674570;
      W_g[13,13] := -0.02423173;
      W_g[13,14] := -0.00389455;
      W_g[13,15] := -0.04698916;
      W_g[13,16] := -0.04386003;
      W_g[13,17] := -0.01447618;
      W_g[13,18] := -0.00030072;
      W_g[13,19] := 0.09379271;
      W_g[13,20] := 0.36890578;
      W_g[13,21] := 0.28695717;
      W_g[13,22] := -0.09331041;
      W_g[13,23] := -0.11805235;
      W_g[13,24] := -0.29436022;
      W_g[13,25] := -0.14414833;
      W_g[13,26] := -0.02907282;
      W_g[13,27] := 0.51352721;
      W_g[13,28] := -0.67788428;
      W_g[13,29] := -0.07989703;
      W_g[13,30] := -0.09920775;
      W_g[13,31] := -0.18299282;
      W_g[13,32] := -0.03875973;
      W_g[13,33] := -0.03526488;
